   REGION Cyclic Error Checks
       IF NOT #Safety_OK_Delayed THEN //11:1
           "Set_Bit_F"(Bit := 0,
                       Bit_Value := 1,
                       Var := #Cnv_Control.Cnv_Errors.Error_Word_1);
       END_IF;

       IF #Cnv_Control.Motor.Error THEN
           "Set_Bit_F"(Bit := 0,
                       Bit_Value := 1,
                       Var := #Cnv_Control.Cnv_Errors.Error_Word_4);
       END_IF;

       IF #Cnv_Control.Instruction.Stop THEN //HMI STOP
           "Set_Bit_F"(Bit := 1,
                       Bit_Value := 1,
                       Var := #Cnv_Control.Cnv_Errors.Error_Word_1);
       END_IF;

       IF #Cnv_Control.Safety_Stop_Cnrl.Error THEN
           "Set_Bit_F"(Bit := 1,
                       Bit_Value := 1,
                       Var := #Cnv_Control.Cnv_Errors.Error_Word_4);
       END_IF;

       // IF ((#ID_Decoded.VTD = 1 AND "Errors_Profinet_1".%X8) OR
       //     (#ID_Decoded.VTD = 2 AND "Errors_Profinet_3".%X7) OR
       //     (*#ID_Decoded.VTD = 3 AND "Errors_Profinet_5".%X4) OR *)
       //     (#ID_Decoded.VTD = 4 AND "Errors_Profinet_7".%X1) OR
       //     (#ID_Decoded.VTD = 5 AND "Errors_Profinet_8".%X6)) AND #Cnv_Control.Mode <> 1
       // THEN //Profinet error
       //     "Set_Bit_F"(Bit := 3,
       //                 Bit_Value := 1,
       //                 Var := #Cnv_Control.Cnv_Errors.Error_Word_3);
       // END_IF;


       // go to error state
       IF #Cnv_Control.Cnv_Errors.Error_Word_1 <> 0 OR
           #Cnv_Control.Cnv_Errors.Error_Word_2 <> 0 OR
           #Cnv_Control.Cnv_Errors.Error_Word_3 <> 0 OR
           #Cnv_Control.Cnv_Errors.Error_Word_4 <> 0
       THEN
           #Cnv_Control.Error := TRUE;
           #State := 400;
       END_IF;
   END_REGION

   REGION VFD
       //Status
       #Cnv_Control.Motor.Ready := (#Cnv_Control.Inputs.VFD_Status.%X0 OR #Cnv_Control.Inputs.VFD_Status.%X1) AND NOT #Cnv_Control.Motor.Error;
       #Cnv_Control.Motor.Error := #Cnv_Control.Inputs.VFD_Status.%X3 OR #Cnv_Control.Inputs.VFD_Status.%X7 OR NOT #Cnv_Control.Inputs.VFD_Status.%X13;
       #Cnv_Control.Motor.Enabled := #Cnv_Control.Inputs.VFD_Status.%X2;
       #Cnv_Control.Motor.Actual_Current := SCALE_X(MIN := 0,
                                                    VALUE := NORM_X(MIN := 0,
                                                                    VALUE := #Cnv_Control.Inputs.VFD_ActualCurrent,
                                                                    MAX := 16384),
                                                    MAX := 1.98);


       //Actual Speed
       IF #MainSetpoint > 0 THEN
           #Cnv_Control.Motor.Speed_Actual := SCALE_X(MIN := 0,
                                                      VALUE := NORM_X(MIN := 0,
                                                                      VALUE := #Cnv_Control.Inputs.VFD_Speed_Actual,
                                                                      MAX := 16384),
                                                      MAX := 130);

           #Cnv_Control.Motor.Actual_Torque := SCALE_X(MIN := 0,
                                                       VALUE := NORM_X(MIN := 0,
                                                                       VALUE := #Cnv_Control.Inputs.VFD_ActualTorque,
                                                                       MAX := 16384),
                                                       MAX := 100);
       ELSIF #MainSetpoint < 0 THEN
           #Cnv_Control.Motor.Speed_Actual := SCALE_X(MIN := 0,
                                                      VALUE := NORM_X(MIN := 0,
                                                                      VALUE := #Cnv_Control.Inputs.VFD_Speed_Actual * -1,
                                                                      MAX := 16384),
                                                      MAX := 130);

           #Cnv_Control.Motor.Actual_Torque := SCALE_X(MIN := 0,
                                                       VALUE := NORM_X(MIN := 0,
                                                                       VALUE := #Cnv_Control.Inputs.VFD_ActualTorque * -1,
                                                                       MAX := 16384),
                                                       MAX := 100);
       ELSE
           #Cnv_Control.Motor.Speed_Actual := 0;
           #Cnv_Control.Motor.Actual_Torque := 0;
       END_IF;

       //MAIN SETPOINT
       IF #Cnv_Control.Motor.Forward THEN
           #MainSetpoint := (SCALE_X(MIN := 0,
                                     VALUE := NORM_X(MIN := 0,
                                                     VALUE := #Cnv_Control.Motor.Speed (** 1.681*),
                                                     MAX := 130),
                                     MAX := 1865.0) * -1);
       ELSIF #Cnv_Control.Motor.Reverse THEN
           #MainSetpoint := SCALE_X(MIN := 0,
                                    VALUE := NORM_X(MIN := 0,
                                                    VALUE := #Cnv_Control.Motor.Speed (** 1.681*),
                                                    MAX := 130),
                                    MAX := 1865.0);
       ELSE
           #MainSetpoint := 0;
       END_IF;

       IF #Safety_OK THEN
           #ConfigAxis := 16#003F;
       ELSE
           #ConfigAxis := 16#003D;
       END_IF;

           #SinaSpeed(EnableAxis := #Cnv_Control.Motor.Forward OR #Cnv_Control.Motor.Reverse,
                      AckError := #Cnv_Control.Instruction.Reset OR "Reset_All" OR #HMI_Reset,
                      SpeedSp := #MainSetpoint,
                      RefSpeed := 1865.0,
                      ConfigAxis := #ConfigAxis,
                      HWIDSTW := #Cnv_Settings.G120_Hardware_ID,
                      HWIDZSW := #Cnv_Settings.G120_Hardware_ID);


   END_REGION

   #HMI_Reset := "Screen_DB_1".Reset_All[1] OR "Screen_DB_1".Reset_All[2] OR "CNV_HMI"."Reset(1)"[1] OR "CNV_HMI"."Reset(1)"[2];
   ;
END_FUNCTION_BLOCK

FUNCTION_BLOCK "Safety_Stops_FB"   // FB7, SCL
{ S7_Optimized_Access := 'TRUE' }
VERSION : 0.1
// stored: AutoNumber true, IsIECCheckEnabled false, IsRetainMemResEnabled false, MemoryReserve 100, SetENOAutomatically false, UDAEnableTagReadback false
   VAR_INPUT
      Sys_No : UInt;
      Mode : UInt;
      Timeout : UInt;
      Reset : Bool;
   END_VAR
   VAR_IN_OUT
      Sfts_Control : "Sfts_Control";
   END_VAR
   VAR
      State : UInt;
      LP_Timer { ExternalAccessible := 'False'; ExternalVisible := 'False'; ExternalWritable := 'False'} : TON_TIME;
      T_Run { S7_SetPoint := 'True'} : TOF_TIME;
      Timer_1 : Time;
   END_VAR
BEGIN
   #Sfts_Control.Enabled := #Sfts_Control.Instruction.Enable := #Mode = 2 OR #Mode = 3;

   //MODES
   IF (#Mode = 1 OR #Mode = 5) AND NOT #Sfts_Control.Error THEN
       #State := 500;
   END_IF;

   (*
   TODO
   1. Need to add the mode and running checks for manual mode
   2. Add output for safety stop brake.

   Mode select is done via the HMI. Might add external mode select switches.

           Mode select mask:
           0: Disabled
           1: Manual
           2: Semi-Auto
           3: Auto
           4: Teach - N/A for Cnv
           5: Maintenance

   Device ID Format: XXYYZZ    
   XX = Device type   
       01   VTD
       10  Cnv_Front_of_VTD
       11  Cnv_Rear_of_VTD
       12  Cnv_On_Extractor
       20  Safety_Stop_Front_of_VTD
       21  Safety_Stop_Rear_of_VTD
   YY = Floor   
   ZZ = VTD Connected to 
   *)


   REGION Cyclic Checks
       //Update variables
       #Sfts_Control.SM_State := #State;

       #LP_Timer(IN := #Sfts_Control.Running,
                 PT := UINT_TO_TIME(#Timeout));

       //STOPPER STATE
       IF #Sfts_Control.Inputs.DP_Extended AND NOT #Sfts_Control.Inputs.DP_Retracted THEN
           #Sfts_Control.LP_State := 1; // EXTENDED
       ELSIF NOT #Sfts_Control.Inputs.DP_Extended AND #Sfts_Control.Inputs.DP_Retracted THEN
           #Sfts_Control.LP_State := 0; //RETRACTED
       ELSE
           #Sfts_Control.LP_State := 2; //LOST
       END_IF;;
   END_REGION

   REGION Auto Mode 
           CASE #State OF
               0: //IDLE MODE
                   IF #Mode = 2 OR #Mode = 3 THEN
                       IF #Sfts_Control.Instruction.Enable AND #Sfts_Control.Error = 0 THEN
                           #Sfts_Control.Enabled := TRUE;
                           #State := 10;
                       END_IF;
                   END_IF;
               10: //Standby
                   IF NOT #Sfts_Control.Running AND #Sfts_Control.Error = 0 AND
                       (#Sfts_Control.Instruction.Extend AND (#Mode = 3 OR #Mode = 2)) OR (#Sfts_Control.Instruction.Manual_Extend AND #Mode = 2) THEN
                       IF #Sfts_Control.Inputs.DP_Extended THEN
                           ; // Complete the task as the LP ar already extended
                       ELSIF #Sfts_Control.Inputs.DP_Retracted THEN
                           #Sfts_Control.Running := True;
                           #State := 20;
                       ELSE
                           #Sfts_Control.Error := 0; //Unknown locking pin state
                           #State := 400;
                       END_IF;
                   ELSIF NOT #Sfts_Control.Running AND #Sfts_Control.Error = 0 AND
                       (#Sfts_Control.Instruction.Retract AND #Mode = 3) OR (#Sfts_Control.Instruction.Manual_Retract AND #Mode = 2) THEN
                       IF #Sfts_Control.Inputs.DP_Retracted THEN
                           ; // Complete the task as the LP ar already extended
                       ELSIF #Sfts_Control.Inputs.DP_Extended THEN
                           #Sfts_Control.Running := True;
                           #State := 40;
                       ELSE
                           #Sfts_Control.Error := 0; //Unknown locking pin state
                           #State := 400;
                       END_IF;
                   END_IF;

               20: //Extend safety locking pins
                   #Sfts_Control.Motor_Extend := TRUE;
                   IF #Sfts_Control.Inputs.DP_Extended THEN
                       #Sfts_Control.Motor_Extend := FALSE;
                       #Sfts_Control.Running := FALSE;
                       #State := 0;
                   END_IF;

               40: //Retract safety locking pins
                   #Sfts_Control.Motor_Retract := TRUE;
                   IF #Sfts_Control.Inputs.DP_Retracted THEN
                       #Sfts_Control.Motor_Retract := FALSE;
                       #Sfts_Control.Running := FALSE;
                       #State := 0;
                   END_IF;

               400: // Error#Sfts_Control
                   #Sfts_Control.Motor_Retract := FALSE;
                   #Sfts_Control.Motor_Extend := FALSE;
                   #Sfts_Control.Running := FALSE;
                   #LP_Timer(IN := FALSE,
                             PT := T#0S);
                   IF #Reset OR "Reset_All" OR
                       "Screen_DB_1".Reset_All[1] OR "Screen_DB_1".Reset_All[2] OR
                       "CNV_HMI"."Reset(1)"[1] OR "CNV_HMI"."Reset(1)"[2]
                   THEN
                       #Sfts_Control.Error := FALSE;
                       #State := 0;
                   END_IF;

               500:
                   IF #Sfts_Control.Instruction.Manual_Extend AND NOT #Sfts_Control.Inputs.DP_Extended THEN
                       #Sfts_Control.Motor_Extend := TRUE;
                       #Sfts_Control.Running := TRUE;
                   ELSIF #Sfts_Control.Instruction.Manual_Retract AND NOT #Sfts_Control.Inputs.DP_Retracted THEN
                       #Sfts_Control.Motor_Retract := TRUE;
                       #Sfts_Control.Running := TRUE;
                   ELSE
                       #Sfts_Control.Motor_Extend := FALSE;
                       #Sfts_Control.Motor_Retract := FALSE;
                       #Sfts_Control.Running := FALSE;
                   END_IF;

                   IF #Mode <> 1 AND #Mode <> 5 THEN
                       #State := 0;
                   END_IF;
           END_CASE;
   END_REGION

   REGION Cyclic Error Checks
       IF #Sfts_Control.Inputs.DP_Extended AND #Sfts_Control.Inputs.DP_Retracted THEN
           #Sfts_Control.Error := TRUE; //Cant have the locking pins extended and retracted at the same time11
       END_IF;

       // Statement section REGION
       IF #LP_Timer.Q THEN
           #Sfts_Control.Error := TRUE;//locking pin timeout
       END_IF;

       IF #Sfts_Control.Error THEN
           #State := 400;
       END_IF;
   END_REGION

   REGION Assign outputs
       #T_Run(IN := #Sfts_Control.Motor_Extend OR #Sfts_Control.Motor_Retract,
                             PT := #Timer_1);

   END_REGION
END_FUNCTION_BLOCK

FUNCTION_BLOCK "Light_Bars"   // FB6, SCL
{ S7_Optimized_Access := 'TRUE' }
VERSION : 0.1
// stored: AutoNumber true, IsIECCheckEnabled false, IsRetainMemResEnabled false, MemoryReserve 100, SetENOAutomatically false, UDAEnableTagReadback false
   VAR_INPUT
      VTD_Mode : UInt;
      VTD_Speed : Int;
      Fault : Bool;
   END_VAR
   VAR_OUTPUT
      Animation_B1 : Byte;
      Color_B1 : Byte;
      Speed_B1 : Byte;
      Animation_B2 : Byte;
      Color_B2 : Byte;
      Speed_B2 : Byte;
   END_VAR
BEGIN
   //Commands for Light Bar

   IF #VTD_Mode = 0 AND NOT #Fault THEN // (0)Disabled = No light  
       #Animation_B1:= #Animation_B2:= 0;

   ELSIF #VTD_Mode = 1 AND #VTD_Speed = 0 AND  NOT #Fault AND NOT "SinaSpeed_VTD_DB_1".EnableAxis THEN // (1)Manual= Yellow Stop
       #Animation_B1 := #Animation_B2 := 1;
       #Color_B1 := #Color_B2 := 4;

   ELSIF #VTD_Mode = 1 AND #VTD_Speed > 0 AND #VTD_Speed <= 33 AND  NOT #Fault AND "SinaSpeed_VTD_DB_1".EnableAxis THEN // (1)Manual= Yellow until 33%
       #Animation_B1 := #Animation_B2 := 2;
       #Speed_B1 := #Speed_B2 := 2;
       #Color_B1 := #Color_B2 := 4;

   ELSIF #VTD_Mode = 1 AND #VTD_Speed > 33 AND #VTD_Speed <= 100 AND  NOT #Fault THEN // (1)Manual= Yellow until 66%
       #Animation_B1 := #Animation_B2 := 2;
       #Speed_B1 := #Speed_B2 := 0;
       #Color_B1 := #Color_B2 := 4;

   // ELSIF #VTD_Mode = 1 AND #VTD_Speed > 66 AND #VTD_Speed <= 100 AND  NOT #Fault THEN // (1)Manual= Yellow until 100%
   //     #Animation_B1 := #Animation_B2 := 2;
   //     #Speed_B1 := #Speed_B2 := 1;
   //     #Color_B1 := #Color_B2 := 4;

   ELSIF #VTD_Mode = 2 AND #VTD_Speed = 0 AND  NOT #Fault AND NOT "SinaSpeed_VTD_DB_1".EnableAxis THEN // (2)Semi-auto = Blue Stop
       #Animation_B1 := #Animation_B2 := 1;
       #Color_B1 := #Color_B2 := 9;
       #Speed_B1 := #Speed_B2 := 0;

   ELSIF #VTD_Mode = 2 AND #VTD_Speed > 0 AND #VTD_Speed <= 33 AND  NOT #Fault AND "SinaSpeed_VTD_DB_1".EnableAxis THEN // (2)Semi-auto = Blue until 33%
       #Animation_B1 := #Animation_B2 := 2;
       #Speed_B1 := #Speed_B2 := 2;
       #Color_B1 := #Color_B2 := 9;

   ELSIF #VTD_Mode = 2 AND #VTD_Speed > 33 AND #VTD_Speed <= 100 AND  NOT #Fault THEN // (2)Semi-auto = Blue until 66%
       #Animation_B1 := #Animation_B2 := 2;
       #Speed_B1 := #Speed_B2 := 0;
       #Color_B1 := #Color_B2 := 9;

   // ELSIF #VTD_Mode = 2 AND #VTD_Speed > 66 AND #VTD_Speed <= 100 AND  NOT #Fault THEN // (2)Semi-auto = Blue until 100%
   //     #Animation_B1 := #Animation_B2 := 2;
   //     #Speed_B1 := #Speed_B2 := 1;
   //     #Color_B1 := #Color_B2 := 9;

   ELSIF #VTD_Mode = 3 AND #VTD_Speed = 0 AND  NOT #Fault AND NOT "SinaSpeed_VTD_DB_1".EnableAxis THEN // (3)Auto = Green Stop
       #Animation_B1 := #Animation_B2 := 1;
       #Color_B1 := #Color_B2 := 0;

   ELSIF #VTD_Mode = 3 AND #VTD_Speed > 0 AND #VTD_Speed <= 33 AND  NOT #Fault AND "SinaSpeed_VTD_DB_1".EnableAxis THEN // (3)Auto = Green until 33%
       #Animation_B1 := #Animation_B2 := 2;
       #Speed_B1 := #Speed_B2 := 2;
       #Color_B1 := #Color_B2 := 0;

   ELSIF #VTD_Mode = 3 AND #VTD_Speed > 33 AND #VTD_Speed <= 100 AND  NOT #Fault THEN // (3)Auto = Green until 66%
       #Animation_B1 := #Animation_B2 := 2;
       #Speed_B1 := #Speed_B2 := 0;
       #Color_B1 := #Color_B2 := 0;

   // ELSIF #VTD_Mode = 3 AND #VTD_Speed > 66 AND #VTD_Speed <= 100 AND  NOT #Fault THEN // (3)Auto = Green until 100%
   //     #Animation_B1 := #Animation_B2 := 2;
   //     #Speed_B1 := #Speed_B2 := 1;
   //     #Color_B1 := #Color_B2 := 0;

   ELSIF #VTD_Mode = 4 AND #VTD_Speed = 0 AND  NOT #Fault THEN // (4)Tech = Orange Stop
       #Animation_B1 := #Animation_B2 := 1;
       #Color_B1 := #Color_B2 := 2;

   ELSIF #VTD_Mode = 4 AND #VTD_Speed > 0 AND #VTD_Speed <= 33 AND  NOT #Fault THEN // (4)Tech = Orange until 33%
       #Animation_B1 := #Animation_B2 := 2;
       #Speed_B1 := #Speed_B2 := 2;
       #Color_B1 := #Color_B2 := 2;

   ELSIF #VTD_Mode = 4 AND #VTD_Speed > 33 AND #VTD_Speed <= 66 AND  NOT #Fault THEN // (4)Tech = Orange until 66%
       #Animation_B1 := #Animation_B2 := 2;
       #Speed_B1 := #Speed_B2 := 0;
       #Color_B1 := #Color_B2 := 2;

   ELSIF #VTD_Mode = 4 AND #VTD_Speed > 66 AND #VTD_Speed <= 100 AND  NOT #Fault THEN // (4)Tech = Orange until 100%
       #Animation_B1 := #Animation_B2 := 2;
       #Speed_B1 := #Speed_B2 := 1;
       #Color_B1 := #Color_B2 := 2;

   ELSIF #VTD_Mode = 5 AND #VTD_Speed = 0 AND  NOT #Fault THEN // (5)Maintenance = White Stop
       #Animation_B1 := #Animation_B2 := 1;
       #Color_B1 := #Color_B2 := 19;

   ELSIF #VTD_Mode = 5 AND #VTD_Speed > 0 AND #VTD_Speed <= 33 AND  NOT #Fault THEN // (5)Maintenance = White until 33%
       #Animation_B1 := #Animation_B2 := 2;
       #Speed_B1 := #Speed_B2 := 2;
       #Color_B1 := #Color_B2 := 19;

   ELSIF #VTD_Mode = 5 AND #VTD_Speed > 33 AND #VTD_Speed <= 66 AND  NOT #Fault THEN // (5)Maintenance = White until 66%
       #Animation_B1 := #Animation_B2 := 2;
       #Speed_B1 := #Speed_B2 := 0;
       #Color_B1 := #Color_B2 := 19;

   ELSIF #VTD_Mode = 5 AND #VTD_Speed > 66 AND #VTD_Speed <= 100 AND  NOT #Fault THEN // (5)Maintenance = White until 100%
       #Animation_B1 := #Animation_B2 := 2;
       #Speed_B1 := #Speed_B2 := 1;
       #Color_B1 := #Color_B2 := 19;

   ELSIF #Fault THEN // Fault = Flash Red
       #Animation_B1:= #Animation_B2 := 2;
       #Color_B1:=#Color_B2 := 1;
   END_IF;
END_FUNCTION_BLOCK

FUNCTION_BLOCK "SICK_Lector_CLV6xx_PNDP"   // FB72, SCL
TITLE = SICK Lector6xx / CLV6xx function block
{ S7_Optimized_Access := 'TRUE' }
AUTHOR : SICKAG
FAMILY : Ident
VERSION : 1.2
// This function block is used for a communication between a SICK Lector6xx / SICK CLV6xx code reader and a Siemens S7-1200/S7-1500 PLC via  PROFINET/PROFIBUS
// stored: AutoNumber false, IsIECCheckEnabled false, IsRetainMemResEnabled false, MemoryReserve 100, SetENOAutomatically false, UDAEnableTagReadback false
   VAR_INPUT
      HWInputIdent : HW_IO;   // Hardware identification number of the input module
      HWInputLength : USInt;   // Size of the input module
      HWOutputIdent : HW_IO;   // Hardware identification number of the output module
      HWOutputLength : USInt;   // Size of the output module
      CANId : USInt;   // CAN ID (0= Master / No CAN network)
      TOut : Time := T#10s;   // Time out
      Req : Bool;   // A positive edge starts the request
      TriggerOn : Bool;   // Select: Trigger On to open the reading gate via a SW-Trigger command
      TriggerOff : Bool;   // Select: Trigger Off to close the reading gate via a SW-Trigger command
      Matchcode : Bool;   // Select: Matchcode (details at #Data)
      SavePermanent : Bool;   // Select: Save permanent
      ComTest : Bool;   // Select: Communication test
      FreeCommand : Bool;   // Select: Free command (details at #Data)
   END_VAR
   VAR_OUTPUT
      RdDone : Bool;   // Positive edge: A reading result sent by the device was received
      ReqDone : Bool;   // Request done
      ReqBusy : Bool;   // Request in process
      Error : Bool;   // Error detected
      Errorcode : DWord;   // Error code (see documentation)
   END_VAR
   VAR_IN_OUT
      Data : "ST_SICK_Lector_CLV6xx";   // Command arguments and result outputs of the FB actions
   END_VAR
   VAR
      bTriggerReq { ExternalAccessible := 'False'; ExternalVisible := 'False'; ExternalWritable := 'False'} : Bool;   // Rising edge detection
      bTriggerReqMem { ExternalAccessible := 'False'; ExternalVisible := 'False'; ExternalWritable := 'False'} : Bool;   // Rising edge detection
      bTriggerDone { ExternalAccessible := 'False'; ExternalVisible := 'False'; ExternalWritable := 'False'} : Bool;   // Rising edge detection
      bTriggerDoneMem { ExternalAccessible := 'False'; ExternalVisible := 'False'; ExternalWritable := 'False'} : Bool;   // Rising edge detection
      bTriggerError { ExternalAccessible := 'False'; ExternalVisible := 'False'; ExternalWritable := 'False'} : Bool;   // Rising edge detection
      bTriggerErrorMem { ExternalAccessible := 'False'; ExternalVisible := 'False'; ExternalWritable := 'False'} : Bool;   // Rising edge detection
      bCanActive { ExternalAccessible := 'False'; ExternalVisible := 'False'; ExternalWritable := 'False'} : Bool;   // CAN-Bus active flag
      bDeviceState { ExternalAccessible := 'False'; ExternalVisible := 'False'; ExternalWritable := 'False'} : Bool;   // Current device state (True= Edit-Mode | False= Run-Mode)
      bEnforceLogout { ExternalAccessible := 'False'; ExternalVisible := 'False'; ExternalWritable := 'False'} : Bool;   // Logout enforced
      bReqBusyMem : Bool;   // Backup variable
      iStep { ExternalAccessible := 'False'; ExternalVisible := 'False'; ExternalWritable := 'False'} : USInt;   // Currrent FB step
      iCommandIndex { ExternalAccessible := 'False'; ExternalVisible := 'False'; ExternalWritable := 'False'} : Int;   // Command index
      iCommandLength { ExternalAccessible := 'False'; ExternalVisible := 'False'; ExternalWritable := 'False'} : UInt;   // Length of the command that should be send
      iRecordSize { ExternalAccessible := 'False'; ExternalVisible := 'False'; ExternalWritable := 'False'} : UInt;   // Length of the record array
      iCommandSize { ExternalAccessible := 'False'; ExternalVisible := 'False'; ExternalWritable := 'False'} : UInt;   // Length of the command array
      iReadingResultSize { ExternalAccessible := 'False'; ExternalVisible := 'False'; ExternalWritable := 'False'} : UInt;   // Length of the reading result array
      iIndex { ExternalAccessible := 'False'; ExternalVisible := 'False'; ExternalWritable := 'False'} : UInt;   // Index variable
      nTempErrorCode { ExternalAccessible := 'False'; ExternalVisible := 'False'; ExternalWritable := 'False'} : DWord;   // Temporarily error code
      nLogoutErrorCode { ExternalAccessible := 'False'; ExternalVisible := 'False'; ExternalWritable := 'False'} : DWord;   // Temporarily error code
      arrSelection { ExternalAccessible := 'False'; ExternalVisible := 'False'; ExternalWritable := 'False'} : Array[0..5] of Bool;   // input bit selection
      arrCommand { ExternalAccessible := 'False'; ExternalVisible := 'False'; ExternalWritable := 'False'} : Array[0..499] of Byte;   // Contains the transmitted CoLa command
      arrRecord { ExternalAccessible := 'False'; ExternalVisible := 'False'; ExternalWritable := 'False'} : Array[0..499] of Byte;   // Contains the received telegram
      fbTimeout { ExternalAccessible := 'False'; ExternalVisible := 'False'; ExternalWritable := 'False'; S7_SetPoint := 'True'} : TON_TIME;   // Instance: Timer on delay (Time out)
      fbCCom { ExternalAccessible := 'False'; ExternalVisible := 'False'; ExternalWritable := 'False'; S7_SetPoint := 'True'} : "SICK_CCOMM_PNDP";   // Instance: CoLa communication block
   END_VAR
   VAR_TEMP
      iTemp1 : Int;   // Temporarily variable
      iTemp2 : UDInt;   // Temporarily variable
      iTemp3 : UDInt;   // Temporarily variable
      nFncValue : DWord;   // Get/Set function value
      nFncErrorCode : Word;   // Get/Set function error code
   END_VAR
BEGIN
   (*===========================================================================================
   Name:   SICK_Lector_CLV6xx_PNDP 
   Author: SICK AG
   =============================================================================================
   Description: 
   This function block is used for a communication between a SICK Lector6xx / SICK CLV6xx
   code reader and a Siemens S7-1200/S7-1500 PLC via PROFINET/PROFIBUS.                         

   =============================================================================================
   Features:        
   - Receive reading results of the device, triggered by a command, fieldbus or by a hardware 
     switch. The content of the result can be modified in the "Output Format" option in the
     SOPAS engineeringtool.                                           
   - Open and close a reading gate (software trigger via command)
   - Set a new Matchcode evaluation condition 
   - Save all device parameters permanent                                                  
   - Communication test
   - Send a free defined CoLa-A telegram and receive the result
   - All commands can also be used in a SICK CAN-Bus network

   =============================================================================================
   Version history:
   Date       | Version | Author  | Remark
   ---------------------------------------------------------------------------------------------
   21/02/2014 | V1.0    | SICK AG | Initial version
   07/08/2014 | V1.1    | SICK AG | Replace R_TRIG function 
   24/10/2017 | V1.2    | SICK AG | Avoid initialization warnings which occurs using TIA V13 or higher
   ============================================================================================*)

   (*===================================== INITIALISATION =====================================*)
   #iRecordSize:= 500;         (*Length of the arrRecord array*)
   #iCommandSize:= 500;        (*Length of the arrCommand array*)
   #iReadingResultSize:= 200;  (*Length of the reading result array*)

   (*Rising edge detection*)
   #bTriggerReq:= #Req AND NOT #bTriggerReqMem;
   #bTriggerReqMem:= #Req;
   #bTriggerDone:= #fbCCom.ReqDone AND NOT #bTriggerDoneMem;
   #bTriggerDoneMem:= #fbCCom.ReqDone;
   #bTriggerError:= #fbCCom.Error AND NOT #bTriggerErrorMem;
   #bTriggerErrorMem:= #fbCCom.Error;

   (*Reset the read done flag every cycle*)
   #RdDone:= false;


   (*===================================== ERROR HANDLING =====================================*)
   (* bDeviceState  |  bEnforceLogout  |  Action
          FALSE     |      FALSE       |  Errorcode = Errorcode from last plc cycle
          FALSE     |      TRUE        |  Errorcode = Logout error
          TRUE      |      FALSE       |  Enforce "Logout" command
          TRUE      |      TRUE        |  Errorcode = Logout not possible + Reason*)
   IF #nTempErrorCode <>16#0000_0000 THEN

     (*Enfore "Logout" command*)
     IF #bDeviceState AND NOT #bEnforceLogout THEN
       #bEnforceLogout:= true;
       #iCommandIndex:= 11;                  (*Logout*)
       #nLogoutErrorCode:= #nTempErrorCode;  (*Save current error code*)
       #nTempErrorCode:= 16#0000_0000;       (*Clear currenr error variable*)
       #iStep:= 4;                           (*Create command*)

     (*Logout can not be ensured*)
     ELSIF #bDeviceState AND #bEnforceLogout THEN
       #Errorcode.%W1:= #nTempErrorCode.%W0;  
       #Errorcode.%W0:= 16#0017;  (*Error: Logout can not be ensured (please check the device state)*)

     (*Errorcode = Errorcode from the last plc cycle or logout error*)
     ELSE
       #Errorcode:= #nTempErrorCode;
     END_IF;

     (*Update FB status*)
     IF #nTempErrorCode <> 16#0000_0000 THEN
       #ReqDone:= false;
       #ReqBusy:= false;
       #bReqBusyMem:= false;
       #Error:= true;
       #nTempErrorCode:= 16#0000_0000;
       #nLogoutErrorCode:= 16#0000_0000;
       #iStep:= 0;
       RETURN;
     END_IF;
   END_IF;

   (*Time out detection*)
   #fbTimeout(IN:= #bReqBusyMem, PT:= #TOut);
   IF #fbTimeout.Q THEN
     #nTempErrorCode:= 16#0000_0010; (*Error: Time out*)
   END_IF;

   (*Check if a device error is detected: 'sFA XX'*)
   IF #bTriggerDone AND ((NOT #bCanActive AND
     #arrRecord[0] = 's' AND
     #arrRecord[1] = 'F' AND
     #arrRecord[2] = 'A') OR (#bCanActive AND
     #arrRecord[0] = 's' AND
     #arrRecord[12] = 'F' AND
     #arrRecord[13] = 'A')) THEN

     (*Get the position of the error code*)
     IF #bCanActive THEN
       #iIndex:= 15;
     ELSE
       #iIndex:= 4;
     END_IF;

     "SICK_GetValue"(iTelegramLength:= INT_TO_UINT(#fbCCom.ReqLength),
                     iValueLength:= 0,
                     nValue=> #nFncValue,
                     nErrorCode=> #nFncErrorCode,
                     iPosition:= #iIndex,
                     arrData:= #arrRecord);

     IF #nFncErrorCode = 16#0000 THEN
       #nTempErrorCode.%W1:= DWORD_TO_WORD(#nFncValue);
       #nTempErrorCode.%W0:= 16#0011; (*Error: Device error*)
     ELSE
       #nTempErrorCode.%W1:= #nFncErrorCode;
       #nTempErrorCode.%W0:= 16#0012; (*Error: SICK_GetValue error*)      
     END_IF;
   END_IF;

   (*Error detected*)
   IF #nTempErrorCode <>16#0000_0000 THEN
     RETURN;
   END_IF;


   (*================================= START REQUEST (STEP 1) =================================*)
   IF NOT #bReqBusyMem AND #bTriggerReq THEN
     #ReqDone:= false;
     #ReqBusy:= true;
     #bReqBusyMem:= true;
     #Error:= false;
     #Errorcode:= 16#0000_0000;
     #bDeviceState:= false;
     #bEnforceLogout:= false;

     (*Save the current bit selection for the job*)
     #arrSelection[0]:= #TriggerOn;
     #arrSelection[1]:= #TriggerOff;
     #arrSelection[2]:= #Matchcode;
     #arrSelection[3]:= #SavePermanent;
     #arrSelection[4]:= #ComTest;
     #arrSelection[5]:= #FreeCommand;

     (*Check CAN-ID*)
     IF #CANId > 63 THEN
       #nTempErrorCode:= 16#0000_0014; (*Error invalid CAN Id*)  
     ELSIF #CANId = 0 THEN
       #bCanActive:= false;
       #iStep:= 3; (*Check parameter input*)
     ELSE
       #bCanActive:= true;
       #iStep:= 2; (*Add CAN identifier*)
     END_IF;
   END_IF;


   (*=============================== ADD CAN IDENTIFIER (STEP 2) ==============================*)
   IF #iStep =2 THEN
     Strg_TO_Chars(Strg:= 's{ 00 01 ', pChars:= 0, Cnt=> #iIndex, Chars:=#arrCommand);

     "SICK_SetValue"(bAddBlank:= false,
                     nValue:= #CANId,
                     arrData=> #arrCommand,
                     nErrorCode=> #nFncErrorCode,
                     iPosition:= #iIndex);
     IF #nFncErrorCode <> 16#0000 THEN
       #nTempErrorCode.%W1:= #nFncErrorCode;
       #nTempErrorCode.%W0:= 16#0013; (*Error: SICK_SetValue error*)
     ELSE
       #arrCommand[#iIndex]:= '}';
       #iStep:= 3; (*Check parameter input*)
     END_IF;
   END_IF;


   (*============================= CHECK PARAMETER INPUT (STEP 3) =============================*)
   IF #iStep =3 THEN
     #iTemp1:= 0; (*Counts up the active bit selection*)

     (*Command: Trigger On*)
     IF #arrSelection[0] THEN
       #iTemp1:= #iTemp1+1;
       #iCommandIndex:= 0; (*Send a "Trigger On" command*)
     END_IF;

     (*Command: Trigger Off*)
     IF #arrSelection[1] THEN
       #iTemp1:= #iTemp1+1;
       #iCommandIndex:= 1; (*Send a "Trigger Off" command*)
     END_IF;

     (*Command: Matchcode*)
     IF #arrSelection[2] THEN
       #iTemp1:= #iTemp1+1;

       IF #Data.Matchcode.sName = '' THEN
         #nTempErrorCode:= 16#0000_0022; (*Error: Matchcode name is empty*)
       ELSIF #Data.Matchcode.nCodeType <='$20' OR #Data.Matchcode.nCodeType > '$7E' THEN
         #nTempErrorCode:= 16#0000_0023; (*Error: Invalid code type*)
       END_IF;

       #iCommandIndex:= 10; (*Send a "Login" command*)
     END_IF;

     (*Command: Save permanent*)
     IF #arrSelection[3] THEN 
       #iTemp1:= #iTemp1+1;
       #iCommandIndex:= 10; (*Send a "Login" command*)  
     END_IF;

     (*Command: Communication test*)
     IF #arrSelection[4] THEN
       #iTemp1:= #iTemp1+1;
       #iCommandIndex:= 4; (*Send a "Comm Test" command*)
     END_IF;

     (*Command: Free command*)
     IF #arrSelection[5] THEN
       #iTemp1:= #iTemp1+1;

       (*Check length*)
       IF #bCanActive THEN
         #iTemp2:= INT_TO_UDINT(LEN(#Data.FreeCommand.sCommand))+11;
       ELSE
         #iTemp2:= INT_TO_UDINT(LEN(#Data.FreeCommand.sCommand));
       END_IF;

       IF (LEN(#Data.FreeCommand.sCommand) <=0) OR (#iTemp2 > #iCommandSize) THEN
         #nTempErrorCode:= 16#0000_0020; (*Error: Invalid free command length*)
       END_IF;

       #iCommandIndex:= 5; (*Send a "Free Command" command*)
     END_IF;

     (*Check bit sum of the command selection*)
     IF #iTemp1 <>1 THEN
       #nTempErrorCode:= 16#0000_0015; (*Error: More than one or no parameter selected*)   
     END_IF;

     (*Check if a error was detected*)
     IF #nTempErrorCode = 16#0000_0000 THEN
       #iStep:= 4; (*Create CoLa command*)
     END_IF;
   END_IF;


   (*============================== CREATE COLA COMMAND (STEP 4) ==============================*)
   IF #iStep =4 THEN
     CASE #iCommandIndex OF

     (*Create "Trigger On" command*)
     0:  IF #bCanActive THEN
           Strg_TO_Chars(Strg:= 'MN mTCgateon', pChars:= 12, Cnt=> #iTemp3, Chars:=#arrCommand);
           #iCommandLength:= UDINT_TO_UINT(#iTemp3)+12;
         ELSE
           Strg_TO_Chars(Strg:= 'sMN mTCgateon', pChars:= 0, Cnt=> #iTemp3, Chars:=#arrCommand);
           #iCommandLength:= UDINT_TO_UINT(#iTemp3);
         END_IF;
         #iStep:= 5; (*Send command*)

     (*Create "Trigger Off" command*)
     1:  IF #bCanActive THEN
           Strg_TO_Chars(Strg:= 'MN mTCgateoff', pChars:= 12, Cnt=> #iTemp3, Chars:=#arrCommand);
           #iCommandLength:= UDINT_TO_UINT(#iTemp3)+12;
         ELSE
           Strg_TO_Chars(Strg:= 'sMN mTCgateoff', pChars:= 0, Cnt=> #iTemp3, Chars:=#arrCommand);
           #iCommandLength:= UDINT_TO_UINT(#iTemp3);
         END_IF;
         #iStep:= 5; (*Send command*)

     (*Create "Matchcode" command*)
     2:  IF #bCanActive THEN
           Strg_TO_Chars(Strg:= 'MN mEVSetMatchCode 00 ', pChars:= 12, Cnt=> #iTemp3, Chars:=#arrCommand);
           #iIndex:= UDINT_TO_UINT(#iTemp3+12);
         ELSE
           Strg_TO_Chars(Strg:= 'sMN mEVSetMatchCode 00 ', pChars:= 0, Cnt=> #iTemp3, Chars:=#arrCommand);
           #iIndex:= UDINT_TO_UINT(#iTemp3);
         END_IF;

         (*Add matchcode name*)
         Strg_TO_Chars(Strg:= CONCAT(IN1:= 'name="', IN2:= #Data.Matchcode.sName), pChars:= #iIndex, Cnt=> #iTemp3, Chars:=#arrCommand);
         #iIndex:= #iIndex+UDINT_TO_UINT(#iTemp3);

         (*Add codeType*)
         Strg_TO_Chars(Strg:= '" codeType="', pChars:= #iIndex, Cnt=> #iTemp3, Chars:=#arrCommand);
         #iIndex:= #iIndex+UDINT_TO_UINT(#iTemp3);
         IF #Data.Matchcode.nCodeType = '*' THEN
           Strg_TO_Chars(Strg:= 'dontCare', pChars:= #iIndex, Cnt=> #iTemp3, Chars:=#arrCommand);
           #iIndex:= #iIndex+UDINT_TO_UINT(#iTemp3);
         ELSE
           #arrCommand[#iIndex]:= #Data.Matchcode.nCodeType;
           #iIndex:= #iIndex+1;
         END_IF;

         (*Add Min/Max length*)
         Strg_TO_Chars(Strg:= '" length="', pChars:= #iIndex, Cnt=> #iTemp3, Chars:=#arrCommand);
         #iIndex:= #iIndex+UDINT_TO_UINT(#iTemp3);
         IF #Data.Matchcode.iMinMaxLength = 0 THEN
           Strg_TO_Chars(Strg:= 'dontCare', pChars:= #iIndex, Cnt=> #iTemp3, Chars:=#arrCommand);
           #iIndex:= #iIndex+UDINT_TO_UINT(#iTemp3);
         ELSE
           #arrCommand[#iIndex]:= ((#Data.Matchcode.iMinMaxLength/100) MOD 10)+16#30;     
           #arrCommand[#iIndex+1]:= ((#Data.Matchcode.iMinMaxLength/10) MOD 10)+16#30;
           #arrCommand[#iIndex+2]:= (#Data.Matchcode.iMinMaxLength MOD 10)+16#30;
           #iIndex:= #iIndex+3;
         END_IF;

         (*Add content*)
         Strg_TO_Chars(Strg:= CONCAT(IN1:= '" content="', IN2:= #Data.Matchcode.sContent), pChars:= #iIndex, Cnt=> #iTemp3, Chars:=#arrCommand);
         #iIndex:= #iIndex+UDINT_TO_UINT(#iTemp3);
         #arrCommand[#iIndex]:= '"';


         (*Overwrite the matchcode length*)
         IF #bCanActive THEN
           #nFncValue:= #iIndex-33;      (*Length of the #Matchcode command*)
           #iCommandLength:= #iIndex+1;  (*Length of the whole CoLa command*)
           #iIndex:= 31;                 (*Startindex of the matchcode length*)
         ELSE
           #nFncValue:= #iIndex-22;      (*Length of the #Matchcode command*)
           #iCommandLength:= #iIndex+1;  (*Length of the whole CoLa command*)
           #iIndex:= 20;                 (*Startindex of the matchcode length*)
         END_IF;

         "SICK_SetValue"(bAddBlank:= false,
                         nValue:= #nFncValue,
                         arrData=> #arrCommand,
                         nErrorCode=> #nFncErrorCode,
                         iPosition:=#iIndex);
         IF #nFncErrorCode <> 16#0000 THEN
           #nTempErrorCode.%W1:= #nFncErrorCode;
           #nTempErrorCode.%W0:= 16#0013; (*Error: SICK_SetValue error*)
         ELSE
           #iStep:= 5; (*Send command*)
         END_IF;

     (*Create "Save Permanent" command*)   
     3:  IF #bCanActive THEN
           Strg_TO_Chars(Strg:= 'MN mEEwriteall', pChars:= 12, Cnt=> #iTemp3, Chars:=#arrCommand);
           #iCommandLength:= UDINT_TO_UINT(#iTemp3+12);
         ELSE
           Strg_TO_Chars(Strg:= 'sMN mEEwriteall', pChars:= 0, Cnt=> #iTemp3, Chars:=#arrCommand);
           #iCommandLength:= UDINT_TO_UINT(#iTemp3);
         END_IF;
         #iStep:= 5; (*Send command*)

     (*Create "Communication Test" command*)
     4:  IF #bCanActive THEN
           Strg_TO_Chars(Strg:= 'RI0', pChars:= 12, Cnt=> #iTemp3, Chars:=#arrCommand);
           #iCommandLength:= UDINT_TO_UINT(#iTemp3)+12;
         ELSE
           Strg_TO_Chars(Strg:= 'sRI0', pChars:= 0, Cnt=> #iTemp3, Chars:=#arrCommand);
           #iCommandLength:= UDINT_TO_UINT(#iTemp3);
         END_IF;
         #iStep:= 5; (*Send command*)

     (*Create "Free Command"*)
     5:  IF #bCanActive THEN
           Strg_TO_Chars(Strg:= DELETE(IN:= #Data.FreeCommand.sCommand, L:=1, P:=1), pChars:= 12, Cnt=> #iTemp3, Chars:=#arrCommand);
           #iCommandLength:= UDINT_TO_UINT(#iTemp3)+12;
         ELSE
           Strg_TO_Chars(Strg:= #Data.FreeCommand.sCommand, pChars:= 0, Cnt=> #iTemp3, Chars:=#arrCommand);
           #iCommandLength:= UDINT_TO_UINT(#iTemp3);
         END_IF;
         #iStep:= 5; (*Send command*)

     (*Create "Login" command*)
     10: IF #bCanActive THEN
           Strg_TO_Chars(Strg:= 'MN SetAccessMode 03 F4724744', pChars:= 12, Cnt=> #iTemp3, Chars:=#arrCommand);
           #iCommandLength:= UDINT_TO_UINT(#iTemp3)+12;
         ELSE
           Strg_TO_Chars(Strg:= 'sMN SetAccessMode 03 F4724744', pChars:= 0, Cnt=> #iTemp3, Chars:=#arrCommand);
           #iCommandLength:= UDINT_TO_UINT(#iTemp3);
         END_IF;
         #iStep:= 5; (*Send command*)

     (*Create "Logout" command*)
     11: IF #bCanActive THEN
           Strg_TO_Chars(Strg:= 'MN Run', pChars:= 12, Cnt=> #iTemp3, Chars:=#arrCommand);
           #iCommandLength:= UDINT_TO_UINT(#iTemp3)+12;
         ELSE
           Strg_TO_Chars(Strg:= 'sMN Run', pChars:= 0, Cnt=> #iTemp3, Chars:=#arrCommand);
           #iCommandLength:= UDINT_TO_UINT(#iTemp3);
         END_IF;
         #iStep:= 5; (*Send command*)

       END_CASE;
   END_IF;


   (*=============================== SEND COLA COMMAND (STEP 5) ===============================*)
   IF #iStep =5 THEN
     IF NOT #fbCCom.ReqBusy AND NOT #bTriggerDone AND NOT #bTriggerError THEN
       #fbCCom.Req:= true;
       #iStep:= 6; (*Wait for the command answer*)
     END_IF;
   END_IF;


   (*========================== WAIT FOR THE COMMAND ANSWER (STEP 6) ==========================*)
   IF #iStep =6 THEN
     (*Communication error*)
     IF #bTriggerError THEN
       #nTempErrorCode:= #fbCCom.Errorcode; (*Error: Communication error*)

       (*Communication done*)
     ELSIF #bTriggerDone THEN
       #iStep:= 7; (*Check the command answer*)
     END_IF;
   END_IF;


   (*============================= CHECK COMMAND RESPONSE (STEP 7) ============================*)
   IF #iStep =7 THEN
     CASE #iCommandIndex OF

     (*Check "Trigger On" response*)
     0:  IF #bCanActive THEN
           IF #arrRecord[0] = 's' AND
             #arrRecord[12] = 'A' AND
             #arrRecord[13] = 'N' AND
             #arrRecord[22] = 'o' AND
             #arrRecord[23] = 'n' AND
             #arrRecord[24] = ' ' AND
             #arrRecord[25] = '1' THEN

             #iStep:= 8; (*Action performed*)
           ELSE
             #nTempErrorCode:= 16#0000_0016; (*Error: Invalid device answer*)                    
           END_IF;
         ELSE
           IF #arrRecord[0] = 's' AND
             #arrRecord[1] = 'A' AND
             #arrRecord[2] = 'N' AND
             #arrRecord[11] = 'o' AND
             #arrRecord[12] = 'n' AND
             #arrRecord[13] = ' ' AND
             #arrRecord[14] = '1' THEN

             #iStep:= 8; (*Action performed*)
           ELSE
             #nTempErrorCode:= 16#0000_0016; (*Error: Invalid device answer*)        
           END_IF;
         END_IF;

     (*Check "Trigger Off" response*)
     1:  IF #bCanActive THEN
           IF #arrRecord[0] = 's' AND
             #arrRecord[12] = 'A' AND
             #arrRecord[13] = 'N' AND
             #arrRecord[22] = 'o' AND
             #arrRecord[23] = 'f' AND
             #arrRecord[24] = 'f' AND
             #arrRecord[25] = ' ' AND
             #arrRecord[26] = '1' THEN

             #iStep:= 8; (*Action performed*)
           ELSE
             #nTempErrorCode:= 16#0000_0016; (*Error: Invalid device answer*)          
           END_IF;
         ELSE
           IF #arrRecord[0] = 's' AND
             #arrRecord[1] = 'A' AND
             #arrRecord[2] = 'N' AND
             #arrRecord[11] = 'o' AND
             #arrRecord[12] = 'f' AND
             #arrRecord[13] = 'f' AND
             #arrRecord[14] = ' ' AND
             #arrRecord[15] = '1' THEN

             #iStep:= 8; (*Action performed*)
           ELSE  
             #nTempErrorCode:= 16#0000_0016; (*Error: Invalid device answer*)          
           END_IF;
         END_IF;

     (*Check "Matchcode" response*)
     2:  IF #bCanActive THEN
           IF NOT(#arrRecord[0] = 's' AND
             #arrRecord[12] = 'A' AND
             #arrRecord[13] = 'N' AND
             #arrRecord[27] = 'o' AND
             #arrRecord[28] = 'd' AND
             #arrRecord[29] = 'e' AND
             #arrRecord[30] = ' ' AND
             #arrRecord[31] = '1') THEN

             #nTempErrorCode:= 16#0000_0016; (*Error: Invalid device answer*)          
           END_IF;
         ELSE
           IF NOT(#arrRecord[0] = 's' AND
             #arrRecord[1] = 'A' AND
             #arrRecord[2] = 'N' AND
             #arrRecord[16] = 'o' AND
             #arrRecord[17] = 'd' AND
             #arrRecord[18] = 'e' AND
             #arrRecord[19] = ' ' AND
             #arrRecord[20] = '1') THEN

             #nTempErrorCode:= 16#0000_0016; (*Error: Invalid device answer*)          
           END_IF;
         END_IF;

         IF #nTempErrorCode = 0 THEN
           #iCommandIndex:= 11; (*Logout*)
           #iStep:= 4;         (*Create command*)
         END_IF;    

     (*Check "Save Permanent" response*)
     3:  IF #bCanActive THEN
           IF NOT(#arrRecord[0] = 's' AND
             #arrRecord[12] = 'A' AND
             #arrRecord[13] = 'N' AND
             #arrRecord[23] = 'a' AND
             #arrRecord[24] = 'l' AND
             #arrRecord[25] = 'l' AND
             #arrRecord[26] = ' ' AND
             #arrRecord[27] = '1') THEN

             #nTempErrorCode:= 16#0000_0016; (*Error: Invalid device answer*)          
           END_IF;
         ELSE
           IF NOT(#arrRecord[0] = 's' AND
             #arrRecord[1] = 'A' AND
             #arrRecord[2] = 'N' AND
             #arrRecord[12] = 'a' AND
             #arrRecord[13] = 'l' AND
             #arrRecord[14] = 'l' AND
             #arrRecord[15] = ' ' AND
             #arrRecord[16] = '1') THEN

             #nTempErrorCode:= 16#0000_0016; (*Error: Invalid device answer*)          
           END_IF;
         END_IF;

         IF #nTempErrorCode = 0 THEN
           #iCommandIndex:= 11; (*Logout*)
           #iStep:= 4;         (*Create command*)
         END_IF;

     (*Check "Communication Test" response*)
     4:  IF #bCanActive THEN
           IF #arrRecord[0] = 's' AND
             #arrRecord[12] = 'R' AND
             #arrRecord[13] = 'A' AND
             #arrRecord[14] = ' ' THEN

             #iStep:= 8; (*Action performed*)
           ELSE
             #nTempErrorCode:= 16#0000_0016; (*Error: Invalid device answer*)          
           END_IF;
         ELSE
           IF #arrRecord[0] = 's' AND
             #arrRecord[1] = 'R' AND
             #arrRecord[2] = 'A' AND
             #arrRecord[3] = ' ' THEN

             #iStep:= 8; (*Action performed*)
           ELSE  
             #nTempErrorCode:= 16#0000_0016; (*Error: Invalid device answer*)          
           END_IF;
         END_IF;

     (*Check "Free command" response*)
     5:  IF #fbCCom.ReqLength <= MAX_LEN(#Data.FreeCommand.sResult) THEN 
           Chars_TO_Strg(Chars:= #arrRecord, pChars:= 0, Cnt:= INT_TO_UINT(#fbCCom.ReqLength),Strg=> #Data.FreeCommand.sResult);
           #iStep:= 8; (*Action performed*)
         ELSE
           #nTempErrorCode:= 16#0000_0021; (*Error: Free command result > Result string*)
         END_IF;

     (*Check "Login" response*)
     10:  IF #bCanActive THEN
           IF NOT(#arrRecord[0] = 's' AND
             #arrRecord[12] = 'A' AND
             #arrRecord[13] = 'N' AND
             #arrRecord[24] = 'M' AND
             #arrRecord[25] = 'o' AND
             #arrRecord[26] = 'd' AND
             #arrRecord[27] = 'e' AND
             #arrRecord[28] = ' ' AND
             #arrRecord[29] = '1') THEN

             #nTempErrorCode:= 16#0000_0016; (*Error: Invalid device answer*)          
           END_IF;
         ELSE
           IF NOT(#arrRecord[0] = 's' AND
             #arrRecord[1] = 'A' AND
             #arrRecord[2] = 'N' AND
             #arrRecord[13] = 'M' AND
             #arrRecord[14] = 'o' AND
             #arrRecord[15] = 'd' AND
             #arrRecord[16] = 'e' AND
             #arrRecord[17] = ' ' AND
             #arrRecord[18] = '1') THEN

             #nTempErrorCode:= 16#0000_0016; (*Error: Invalid device answer*)          
           END_IF;
         END_IF;

         IF #nTempErrorCode = 0 THEN
           IF #arrSelection[2] THEN
             #iCommandIndex:= 2; (*Matchcode*)
             #iStep:= 4;         (*Create command*)
           ELSIF #arrSelection[3] THEN
             #iCommandIndex:= 3; (*Save permanent*)
             #iStep:= 4;         (*Create command*)       
           END_IF;
           #bDeviceState:= true; (*Edit-Mode active*)
         END_IF;

     (*Check "Logout" response*)
     11:  IF #bCanActive THEN
           IF #arrRecord[0] = 's' AND
             #arrRecord[12] = 'A' AND
             #arrRecord[13] = 'N' AND
             #arrRecord[14] = ' ' AND
             #arrRecord[15] = 'R' AND
             #arrRecord[16] = 'u' AND
             #arrRecord[17] = 'n' AND
             #arrRecord[18] = ' ' AND
             #arrRecord[19] = '1' THEN

             #bDeviceState:= false; (*Run-Mode active*)
             #iStep:= 8; (*Action performed*)
           ELSE
             #nTempErrorCode:= 16#0000_0016; (*Error: Invalid device answer*)          
           END_IF;
         ELSE
           IF #arrRecord[0] = 's' AND
             #arrRecord[1] = 'A' AND
             #arrRecord[2] = 'N' AND
             #arrRecord[3] = ' ' AND
             #arrRecord[4] = 'R' AND
             #arrRecord[5] = 'u' AND
             #arrRecord[6] = 'n' AND
             #arrRecord[7] = ' ' AND
             #arrRecord[8] = '1' THEN

             #bDeviceState:= false; (*Run-Mode active*)
             #iStep:= 8; (*Action performed*)
           ELSE  
             #nTempErrorCode:= 16#0000_0016; (*Error: Invalid device answer*)          
           END_IF;
         END_IF;
     END_CASE;
   END_IF;


   (*================================ ACTION PERFORMED (STEP 8) ===============================*)
   IF #iStep =8 THEN
     IF #bEnforceLogout THEN
       #nTempErrorCode:= #nLogoutErrorCode;
     ELSE
       #ReqDone:= true;
       #ReqBusy:= false;
       #bReqBusyMem:= false;
       #iStep:= 0;
     END_IF;
   END_IF;


   (*====================================== COMMUNICATION =====================================*)
   #fbCCom(HWInputIdent:= #HWInputIdent,
           HWInputLength:= #HWInputLength,
           HWOutputIdent:= #HWOutputIdent,
           HWOutputLength:= #HWOutputLength,
           TOut:= #TOut+T#1s,
           CommandLength:= #iCommandLength,
           arrCommand:= #arrCommand,
           arrRecord:= #arrRecord);

   (*Reset the request flag every cycle*)
   #fbCCom.Req:= false;

   (*Read result error*)
   IF #fbCCom.RdLength <0 AND #fbCCom.RdDone THEN
     #Data.ReadingResult.iLength:= -1; (*Error: Reading result longer than record array*)
     FOR #iTemp1:= 1 TO UINT_TO_INT(#iReadingResultSize) DO
       #Data.ReadingResult.arrResult[#iTemp1]:= 16#00;
     END_FOR;

   (*Handling of the reading result*)
   ELSIF #fbCCom.RdDone THEN
     IF #fbCCom.RdLength > #iReadingResultSize THEN
       #Data.ReadingResult.iLength:= -1; (*Error: Reading result longer than reading result array*)
       FOR #iTemp1:= 1 TO UINT_TO_INT(#iReadingResultSize) DO
         #Data.ReadingResult.arrResult[#iTemp1]:= 16#00;
       END_FOR;
     ELSE
       MOVE_BLK(IN:= #arrRecord[0], COUNT:= INT_TO_UINT(#fbCCom.RdLength), OUT=> #Data.ReadingResult.arrResult[1]);
       IF (#Data.ReadingResult.iCounter >=255) THEN
         #Data.ReadingResult.iCounter:= 0;
       ELSE
         #Data.ReadingResult.iCounter:= #Data.ReadingResult.iCounter+1;
       END_IF;
       #Data.ReadingResult.iLength:= #fbCCom.RdLength;
       #RdDone:= true;
     END_IF;
   END_IF;
END_FUNCTION_BLOCK

FUNCTION_BLOCK "SICK_CCOMM_PNDP"   // FB10, SCL
TITLE = SICK_CCOM_PNDP
{ S7_Optimized_Access := 'TRUE' }
AUTHOR : SICKAG
FAMILY : Ident
VERSION : 1.2
// The function block use a Profinet/Probibus connection to communicate with a SICK AutoIdent
// device. The FB makes it possible to send and receive sensor data. The Confirmed Messaging 
// protocol (CM-Protocol) is used to receive even long fragmented read results.
// stored: AutoNumber false, IsIECCheckEnabled false, IsRetainMemResEnabled false, MemoryReserve 100, SetENOAutomatically false, UDAEnableTagReadback false
   VAR_INPUT
      HWInputIdent : HW_IO;   // Hardware identification number of the input module
      HWInputLength : USInt;   // Size of the input module
      HWOutputIdent : HW_IO;   // Hardware identification number of the output module
      HWOutputLength : USInt;   // Size of the output module
      TOut : Time := T#5s;   // Time out
      Req : Bool;   // A positive edge starts the request
      CommandLength : UInt;   // Byte length of the command
   END_VAR
   VAR_OUTPUT
      RdDone : Bool;   // Reading result arrived
      RdLength : Int;   // Byte length of the reading result
      ReqDone : Bool;   // Requested data available
      ReqBusy : Bool;   // Request busy
      ReqLength : Int;   // Byte length of the requested data
      Error : Bool;   // Error
      Errorcode : DWord;   // Error code
   END_VAR
   VAR_IN_OUT
      arrCommand : Array[0..499] of Byte;
      arrRecord : Array[0..499] of Byte;
   END_VAR
   VAR
      bTriggerReq { ExternalAccessible := 'False'; ExternalVisible := 'False'; ExternalWritable := 'False'} : Bool := false;   // Rising edge detection
      bTriggerReqMem { ExternalAccessible := 'False'; ExternalVisible := 'False'; ExternalWritable := 'False'} : Bool := false;   // Rising edge detection
      bReadFrag { ExternalAccessible := 'False'; ExternalVisible := 'False'; ExternalWritable := 'False'} : Bool;
      bWriteFrag { ExternalAccessible := 'False'; ExternalVisible := 'False'; ExternalWritable := 'False'} : Bool;
      bReqBusyMem : Bool;
      iReadStep { ExternalAccessible := 'False'; ExternalVisible := 'False'; ExternalWritable := 'False'} : USInt;
      iWriteStep { ExternalAccessible := 'False'; ExternalVisible := 'False'; ExternalWritable := 'False'} : USInt;
      iReadIndex { ExternalAccessible := 'False'; ExternalVisible := 'False'; ExternalWritable := 'False'} : UInt;
      iWriteIndex { ExternalAccessible := 'False'; ExternalVisible := 'False'; ExternalWritable := 'False'} : UInt;
      iReadHeaderLength { ExternalAccessible := 'False'; ExternalVisible := 'False'; ExternalWritable := 'False'} : UInt;
      iWriteHeaderLength { ExternalAccessible := 'False'; ExternalVisible := 'False'; ExternalWritable := 'False'} : UInt;
      iReadFragmentLength { ExternalAccessible := 'False'; ExternalVisible := 'False'; ExternalWritable := 'False'} : UInt;
      iWriteFragmentLength { ExternalAccessible := 'False'; ExternalVisible := 'False'; ExternalWritable := 'False'} : UInt;
      iRecordSize { ExternalAccessible := 'False'; ExternalVisible := 'False'; ExternalWritable := 'False'} : UInt;
      iCommandSize { ExternalAccessible := 'False'; ExternalVisible := 'False'; ExternalWritable := 'False'} : UInt;
      nTempErrorCode { ExternalAccessible := 'False'; ExternalVisible := 'False'; ExternalWritable := 'False'} : DWord;
      arrInputImage : Array[0..127] of Byte;
      arrOutputImage : Array[0..127] of Byte;
      fbTimeout { ExternalAccessible := 'False'; ExternalVisible := 'False'; ExternalWritable := 'False'; S7_SetPoint := 'True'} : TON_TIME;
   END_VAR
   VAR_TEMP
      iTemp1 : Int;
      iTemp2 : UDInt;
      iTemp3 : UDInt;
   END_VAR
BEGIN
   (*===========================================================================================
   Name:   SICK_CCOMM_PNDP
   Author: SICK AG
   =============================================================================================
   Description: 
   The function block use a Profinet/Probibus connection to communicate with a SICK AutoIdent
   device. The FB makes it possible to send and receive sensor data. The Confirmed Messaging 
   protocol (CM-Protocol) is used to receive even long fragmented read results.

   Send a command:
   The "Req" parameter must be triggered with a rising edge (signal change FALSE to TRUE) in 
   order to carry out the function. For the time during which a valid response has yet to be 
   received from the device, the "ReqBusy" parameter is used to signal  that a response is still 
   pending. The module signals the "ReqDone" = TRUE output parameter when the function has been 
   successfully completed. If data was requested by the device, this data is copied into the 
   Record (arrRecord). The "ReqDone" indicates that new data has been received  for a PLC cycle.
   Only one CoLa-A command request can be send to the same device at one time. 

   Receive a reading result:
   Data sent via trigger command or directly by the device (e.g., direct trigger via a light 
   barrier) is stored in the Record (arrRecord). The "RdDone" output indicates that new data 
   has been received for a PLC cycle. The data sent by the device can be changed or adapted in 
   output format of SOPAS-ET. 

   This AOI supports the folowing SICK devices:
   - Lector6xx
   - RFU6xx
   - CLV6xx 
   - RFH6xx
   =============================================================================================
   Confirmed Messaging Protocol definitions:
   arrInputImage[0]        = Status byte 
   arrInputImage[1]        = Receive counter
   arrInputImage[2]        = Transmit counter back
   arrInputImage[3]        = Command length LSB
   arrInputImage[4]        = Command length MSB
   arrInputImage[5..127]   = Device response (CoLa-A)

   arrOutputImage[0]       = Status byte 
   arrOutputImage[1]       = Receive counter back
   arrOutputImage[2]       = Transmit counter
   arrOutputImage[3]       = Command length LSB
   arrOutputImage[4]       = Command length MSB
   arrOutputImage[5..127]  = Device request (CoLa-A)
   =============================================================================================
   Version history:
   Date       | Version | Created under               | Author  | Remark
   ---------------------------------------------------------------------------------------------
   16/01/2014 | V1.0    | TIA Portal V12 SP1 Update 2 | SICK AG | Initial version
   07/08/2014 | V1.1    | TIA Portal V12 SP1 Update 4 | SICK AG | Replace R_TRIG function 
   22/04/2015 | V1.2    | TIA Portal V12 SP1 Update 4 | SICK AG | Avoid warnings that occur with 
                                                                  TIA V13
   ============================================================================================*)

   (*===================================== INITIALISATION =====================================*)
   #iRecordSize:= 500;   (*Length of the arrRecord array*)
   #iCommandSize:= 500;  (*Length of the arrCommand array*)

   #RdDone:= false;
   #iReadStep:= 0;

   (*Rising edge detection of the request flag*)
   #bTriggerReq:= #Req AND NOT #bTriggerReqMem;
   #bTriggerReqMem:= #Req;

   (*Error detection*)
   IF #nTempErrorCode <>16#0000_0000 THEN
     #ReqDone:= false;
     #ReqBusy:= false;
     #bReqBusyMem:= false;
     #Error:= true;
     #Errorcode:= #nTempErrorCode;
     #nTempErrorCode:= 16#0000_0000;
     #ReqLength:= 0;
     #iWriteStep:= 0;
     RETURN;
   END_IF;

   (*Time out detection*)
   #fbTimeout(IN:=#bReqBusyMem, PT:=#TOut);
   IF #fbTimeout.Q THEN
     #nTempErrorCode:= 16#0000_0001; (*Error: Time out*) 
   END_IF;

   (*Check the hardware ident length of the input module*)
   IF #HWInputLength <8 OR #HWInputLength >128 THEN
     #nTempErrorCode:= 16#0000_0002; (*Error: Incorrect module input length*)
   END_IF;

   (*Check the hardware ident length of the output module*)
   IF #HWOutputLength <8 OR #HWOutputLength >128 THEN
     #nTempErrorCode:= 16#0000_0003; (*Error: Incorrect module output length*)
   END_IF;

   (*Error detected*)
   IF #nTempErrorCode <>16#0000_0000 THEN
     RETURN;
   END_IF;


   (*===================================== COMMUNICATION ======================================*)
   (*Set output data*)
   #iTemp1:= DPWR_DAT(LADDR:= #HWOutputIdent, RECORD:= #arrOutputImage);
   IF #iTemp1 <>0 THEN
     #nTempErrorCode.%W1:= #iTemp1;
     #nTempErrorCode.%W0:= 16#0004; (*Error: Set output data via DPWR_DAT*)
     RETURN;
   END_IF;

   (*Get input data*)
   #iTemp1:= DPRD_DAT(LADDR:= #HWInputIdent, RECORD=> #arrInputImage);
   IF #iTemp1 <>0 THEN
     #nTempErrorCode.%W1:= #iTemp1;
     #nTempErrorCode.%W0:= 16#0005; (*Error: Get input data via DPRD_DAT*)
     RETURN;
   END_IF;

   (*Receive counter ==0 && Receive counter back <>0*)
   IF #arrInputImage[1] =0 AND #arrOutputImage[1] <>0 THEN
     #arrOutputImage[1]:= #arrInputImage[1]; (*Recive counter => Receive counter back*)
     RETURN;
   END_IF;

   (*Transmit counter <> Transmit counter back*)
   IF NOT #bReqBusyMem AND (#arrInputImage[2] <> #arrOutputImage[2]) THEN
     #arrOutputImage[2]:= 0; (*0 => Transmit counter*)
     RETURN;
   END_IF;


   (*============================== HANDLING OF THE RECEIVED DATA =============================*)
   (*New telegram available*)
   IF NOT (#arrInputImage[1] = #arrOutputImage[1]) THEN

     (*Reset error every incoming telegram (Read only mode, e.g. for hand held scanners)*)
     IF #CommandLength <=0 THEN
       #Error:= false;
       #Errorcode:= 16#0000_0000;
     END_IF;

     (*Confirm the receive counter*)
     #arrOutputImage[1]:= #arrInputImage[1];

     (*Get telegram length from the received header*)
     #iReadHeaderLength.%B0:= #arrInputImage[3];
     #iReadHeaderLength.%B1:= #arrInputImage[4];

     (*Check if fragmentation is not active at the moment*)
     IF NOT #bReadFrag THEN
       #iReadIndex:= 0;

       (*Check if fragmentation is needed*)
       IF (#HWInputLength-5) < #iReadHeaderLength THEN
         #bReadFrag:= true;
       END_IF;
     END_IF;

     (*Fragmentation is needed*)
     IF #bReadFrag THEN
       IF (#HWInputLength-5) < #iReadHeaderLength THEN
         #iReadFragmentLength:= #HWInputLength-5;
       ELSE
         #iReadFragmentLength:= #iReadHeaderLength;
       END_IF;

     (*No fragmentation needed*)
     ELSE
       #iReadFragmentLength:= #iReadHeaderLength;
     END_IF;

     (*Copy input data into the output record*)
     IF (#iReadIndex+#iReadFragmentLength) <= #iRecordSize THEN
       MOVE_BLK(IN:= #arrInputImage[5], COUNT:= #iReadFragmentLength, OUT=> #arrRecord[#iReadIndex]);
     END_IF;

     (*Check if all data has been received*)
     IF (#HWInputLength-5) < #iReadHeaderLength THEN
       #iReadIndex:= #iReadIndex+#iReadFragmentLength;

     (*All data has been received*)
     ELSE
       #bReadFrag:= false;
       #iReadStep:= 1;
     END_IF;

     (*Incoming data filter*)
     (* - Check if the receiving telegram os a CoLa answer on a requested 
          comand or a reading result.

         sRA  sWA  sMA  sAN  sAI  sEA  sPX  s{   sSI  sSN  sFA
     sRN  X                                       X    X    X
     sRI  X                                       X    X    X
     sWN       X                                  X    X    X
     sWI       X                                  X    X    X
     sMN            X    X                        X    X    X
     sMI            X         X                   X    X    X
     sEN                           X              X    X    X
     sEI                           X              X    X    X
     sPE                                X         X    X    X
     s{                                      X    X    X    X
     *)
     IF #iReadStep =1 THEN
       (*Filter is only active, while requested data expected*)
       IF #bReqBusyMem THEN
         IF #CommandLength >3 THEN
           (*Get the prefix from the requested command (e.g. 'sRN '*)   
           #iTemp2.%B3:= #arrCommand[0];
           #iTemp2.%B2:= #arrCommand[1];
           #iTemp2.%B1:= #arrCommand[2];
           #iTemp2.%B0:= 16#20;

           (*Get the prefix from the command response (e.g. 'sRA ')*)
           #iTemp3.%B3:= #arrRecord[0];
           #iTemp3.%B2:= #arrRecord[1];
           #iTemp3.%B1:= #arrRecord[2];
           #iTemp3.%B0:= 16#20;
         ELSE
           #iTemp2:= 16#0000_0000;
           #iTemp3:= 16#0000_0000;
         END_IF;

         CASE #iTemp3 OF
         (*'s{  '*)
         16#737B2020:  IF #iTemp2 = 16#737B2020 THEN
                         #iReadStep:= 2; (*Command response*)
                       ELSE
                         #iReadStep:= 3; (*Reading result*)
                       END_IF;

         (*'sRA '*)
         16#73524120:  IF (#iTemp2 = 16#73524E20) OR (#iTemp2 = 16#73524920) THEN
                         #iReadStep:= 2; (*Command response*)
                       ELSE
                         #iReadStep:= 3; (*Reading result*)
                       END_IF;

         (*'sWA '*)
         16#73574120:  IF (#iTemp2 = 16#73574E20) OR (#iTemp2 = 16#73574920) THEN
                         #iReadStep:= 2; (*Command response*)
                       ELSE
                         #iReadStep:= 3; (*Reading result*)
                       END_IF;

         (*'sMA '*)
         16#734D4120:  IF (#iTemp2 = 16#734D4E20) OR (#iTemp2 = 16#734D4920) THEN
                         #iReadStep:= 2; (*Command response*)
                       ELSE
                         #iReadStep:= 3; (*Reading result*)
                       END_IF;

         (*'sAN '*)
         16#73414E20:  IF #iTemp2 = 16#734D4E20 THEN
                         #iReadStep:= 2; (*Command response*)
                       ELSE
                         #iReadStep:= 3; (*Reading result*)
                       END_IF;

         (*'sAI '*)
         16#73414920:  IF #iTemp2 = 16#734D4920 THEN
                         #iReadStep:= 2; (*Command response*)
                       ELSE
                         #iReadStep:= 3; (*Reading result*)
                       END_IF;

         (*'sEA '*)
         16#73454120:  IF (#iTemp2 = 16#73454E20) OR (#iTemp2 = 16#73454920) THEN
                         #iReadStep:= 2; (*Command response*)
                       ELSE
                         #iReadStep:= 3; (*Reading result*)
                       END_IF;

         (*'sPX '*)
         16#73505820:  IF #iTemp2 = 16#73504520 THEN
                         #iReadStep:= 2; (*Command response*)
                       ELSE
                         #iReadStep:= 3; (*Reading result*)
                       END_IF;

         (*'sSI '*)
         16#73534920:  #iReadStep:= 3; (*Reading result*)

         (*'sSN '*)
         16#73534E20:  #iReadStep:= 3; (*Reading result*)

         (*'sFA '*)
         16#73464120:  #iReadStep:= 2; (*Command response*)

         (*Invalid CoLa-A answer*)
         ELSE
           (*Check if a user defined command is used (Request == Response)*)
           FOR #iTemp1:= 0 TO UINT_TO_INT(#CommandLength-1) DO
             IF #arrCommand[#iTemp1] = #arrRecord[#iTemp1] THEN
               #iReadStep:= 2; (*Command response*)
             ELSE
               #iReadStep:= 3; (*Reading result*)
               EXIT;
             END_IF;
           END_FOR;
         END_CASE;

       (*Reading result*)
       ELSE
         #iReadStep:= 3;  (*Reading result*)
       END_IF;
     END_IF;

     (*Incoming telegram is a command response*)
     IF #iReadStep =2 THEN
       IF (#iReadIndex+#iReadFragmentLength) <= #iRecordSize THEN
         #ReqLength:= UDINT_TO_INT(#iReadIndex+#iReadFragmentLength);
         #ReqDone:= true;
         #ReqBusy:= false;
         #bReqBusyMem:= false;
       ELSE
         #nTempErrorCode:= 16#0000_0006; (*Error: Incoming command response > Record size*)
       END_IF;
     END_IF;

     (*Incoming telegram is a reading result*)
     IF #iReadStep =3 THEN
       IF (#iReadIndex+#iReadFragmentLength) <= #iRecordSize THEN
         #RdLength:= UDINT_TO_INT(#iReadIndex+#iReadFragmentLength);
         #RdDone:= true;
       ELSE
         #RdLength:= -1;
         #RdDone:= false;    
       END_IF;
     END_IF;
   END_IF;


   (*=========================== HANDLING OF THE DATA TO BE WRITTEN ===========================*)
   IF #bTriggerReq AND NOT #bReqBusyMem THEN
     #ReqDone:= false;
     #ReqBusy:= true;
     #bReqBusyMem:= true;
     #Error:= false;
     #Errorcode:= 16#0000_0000;
     #iWriteIndex:= 0;

     (*Check command length*)
     IF #CommandLength <=0 THEN
       #nTempErrorCode:= 16#0000_0007; (*Error: Command length <= 0*)
       RETURN;
     ELSIF #CommandLength > #iCommandSize THEN
       #nTempErrorCode:= 16#0000_0008; (*Error: Command length > command array*)
       RETURN;
     END_IF;

     (*Check if the the command telegram must be fragmented*)
     IF (#HWOutputLength-5) < #CommandLength THEN
       #iWriteFragmentLength:= #HWOutputLength-5;
     ELSE
       #iWriteFragmentLength:= #CommandLength;
     END_IF;

     #iWriteHeaderLength:= #CommandLength;
     #iWriteStep:= 1;  
   END_IF;

   (*Write step 1: Command transfer*)
   IF (#iWriteStep =1) AND(#arrInputImage[2] = #arrOutputImage[2]) THEN

     (*Copy command data into the output record*)
     IF((#iWriteIndex+#iWriteFragmentLength) <= #iCommandSize) AND (#iWriteFragmentLength <= (#HWOutputLength-5)) THEN
       MOVE_BLK(IN:= #arrCommand[#iWriteIndex], COUNT:= #iWriteFragmentLength, OUT=> #arrOutputImage[5]);
       (*Increment transmit counter*)
       IF #arrOutputImage[2] = 16#FF THEN
         #arrOutputImage[2]:= 16#01; (*Counter overflow, zero is skipped*)
       ELSE
         #arrOutputImage[2]:= #arrOutputImage[2]+1;
       END_IF;

       (*Set command/fragment length*)
       #arrOutputImage[3]:= #iWriteHeaderLength.%B0;
       #arrOutputImage[4]:= #iWriteHeaderLength.%B1;

       (*Next step*)
       #iWriteStep:= 2;
     ELSE
       #nTempErrorCode:= 16#0000_0009; (*Error: Fragmentation error*)
     END_IF;
       RETURN;
   END_IF;

   (*Write step 2: Fragmentation handling*)
   IF #iWriteStep =2 THEN

     (*Fragmentation is needed*)
     IF (#HWOutputLength-5) < #iWriteHeaderLength THEN
       #bWriteFrag:= true;

       (*Next index*)
       #iWriteIndex:= #iWriteIndex+#iWriteFragmentLength;

       (*Set next header length*)
       #iWriteHeaderLength:= #iWriteHeaderLength-#iWriteFragmentLength;

       (*Set next fragment length*)
       IF (#HWOutputLength-5) < #iWriteHeaderLength THEN
         #iWriteFragmentLength:= #HWOutputLength-5;
       ELSE
         #iWriteFragmentLength:= #iWriteHeaderLength;
       END_IF;

     (*Fragmentation is not needed*)
     ELSE
       #bWriteFrag:= false;
     END_IF;

     (*Next step*)
     #iWriteStep:= 3;
   END_IF;

   (*Write step 3: Check if the transmission of the command/fragment is done*)
   IF #iWriteStep =3 THEN

     (*Transmit counter back == Transmit counter*)
     IF #arrInputImage[2] = #arrOutputImage[2] THEN
       IF #bWriteFrag THEN
         #iWriteStep:= 1;
       ELSE
         #iWriteStep:= 0;
       END_IF;
     END_IF;
   END_IF;
END_FUNCTION_BLOCK

FUNCTION_BLOCK "SICK_Lector_Control_FB"   // FB19, SCL
{ S7_Optimized_Access := 'TRUE' }
VERSION : 0.1
// stored: AutoNumber true, IsIECCheckEnabled false, IsRetainMemResEnabled false, MemoryReserve 100, SetENOAutomatically false, UDAEnableTagReadback false
   VAR_INPUT
      Rd_Done : Bool;
      Req_Done : Bool;
      Req_Busy : Bool;
      Error : Bool;
      arrResult : Array[1..200] of Byte;
      iCounter : USInt;
      iLength : Int;
      Error_Code : DWord;
   END_VAR
   VAR_OUTPUT
      Test_Comm : Bool;
      Enable_Trigger : Bool;
      Disable_Trigger : Bool;
      Enable_Req : Bool;
      Result : String;
      Test_OK : Bool;
   END_VAR
   VAR_IN_OUT
      Test_Comm_HMI : Bool;
      Enable_HMI : Bool;
      Disable_HMI : Bool;
      Auto_Start_Lector : Bool;
      Auto_Stop_Lector : Bool;
   END_VAR
   VAR
      "Timer" { S7_SetPoint := 'True'} : TON_TIME;
      R_Done_DB { S7_SetPoint := 'True'} : R_TRIG;
      T_Reset_DB { S7_SetPoint := 'True'} : TON_TIME;
   END_VAR
BEGIN
   //Communication Test
   IF #Test_Comm_HMI THEN
       #Test_Comm := 1;
       #Enable_Req := 1;
       #Timer.TON(IN:=True,
                              PT:=t#1s);
   END_IF;

   //TEST OK
   IF #Req_Done AND #Timer.Q AND NOT #Error THEN
       #Test_OK := 1;
       #Test_Comm := 0;
       #Enable_Req := 0;
       #Test_Comm_HMI := 0;
       #Timer.TON(IN := FALSE,
                              PT := t#0s);
   END_IF;

   //ERROR
   IF #Timer.Q AND #Error THEN
           #Test_OK := 0;
           #Test_Comm := 0;
           #Enable_Req := 0;
           #Test_Comm_HMI := 0;
           #Timer.TON(IN := FALSE,
                                  PT := t#0s);
       END_IF;

   //Enable Trigger
       IF #Enable_HMI OR #Auto_Start_Lector THEN
       #Enable_Trigger := 1;
       #Enable_Req := 1;
       #Disable_HMI := 0;
       #Disable_Trigger := 0;
   //Disable Trigger
   ELSIF #Disable_HMI OR #"Auto_Stop_Lector" THEN
       #Disable_Trigger := 1;
       #Enable_Req := 1;
       #Enable_HMI := 0;
       #Enable_Trigger := 0;
   ELSE
       #Enable_Trigger := 0;
       #Enable_Req := 0;
       #Disable_Trigger := 0;
   END_IF;


   #R_Done_DB(CLK:=#Rd_Done);

   IF #R_Done_DB.Q OR #T_Reset_DB.Q OR
       (#Enable_HMI AND #Disable_HMI)
   THEN
       #Disable_HMI := 0;
       #Enable_Trigger := 0;
       #Disable_Trigger := 0;
       #Enable_Req := 0;
       #T_Reset_DB.TON(IN := FALSE,
                               PT := T#0S);
               #Auto_Stop_Lector := 0;
   END_IF;

   #T_Reset_DB(IN:=(#Enable_HMI OR #Disable_HMI OR #Auto_Start_Lector OR #Auto_Stop_Lector),
                 PT:=T#10S);


   #Result := "ByteArrayToString_1"(Lenght := #iLength, ByteArray := #arrResult);
END_FUNCTION_BLOCK

FUNCTION_BLOCK "Barcode_Station_FB"   // FB33, SCL
{ S7_Optimized_Access := 'TRUE' }
VERSION : 0.1
// stored: AutoNumber true, IsIECCheckEnabled false, IsRetainMemResEnabled false, MemoryReserve 100, SetENOAutomatically false, UDAEnableTagReadback false
   VAR_INPUT
      Sick_Result : String;
   END_VAR
   VAR_OUTPUT
      "Counter" : UInt;
   END_VAR
   VAR_IN_OUT
      Station_Control : "Barcode_Station_UDT";
      Auto_Start_Lector : Bool;
      Auto_Stop_Lector : Bool;
   END_VAR
   VAR
      State : UInt;
      R_Start_DB { S7_SetPoint := 'True'} : R_TRIG;
      T_Read_DB { S7_SetPoint := 'True'} : TON_TIME;
   END_VAR
   VAR_TEMP
      StartPos : Int;
      EndPos : Int;
      Code : String;
   END_VAR
BEGIN
   #R_Start_DB(CLK := #Station_Control.Start);

   IF #R_Start_DB.Q THEN
       IF #State = 0 THEN
           #State := 10;
       END_IF;
   END_IF;

   CASE #State OF
       0: // IDLE
           #Station_Control.Running := FALSE;
           #Station_Control.Ready := TRUE;
           #T_Read_DB(IN := FALSE,
                      PT := T#0S);

       10: // Start
           #Station_Control.Barcode := '';
           #Station_Control.Done := FALSE;
           #Station_Control.Valid := FALSE;
           #Station_Control.Ready := FALSE;
           #Station_Control.Running := TRUE;
           #State := 20;

       20: // Reading code
           #Station_Control.Start := FALSE;
           #Station_Control."Reading Gate number" := "FindStringField"(FieldName := 'Number', JsonStr := #Sick_Result);
           #Station_Control.Barcode := "FindStringField"(FieldName := 'Code', JsonStr := #Sick_Result);
           #Station_Control."Number of Reading Gates" := "FindStringField"(FieldName := 'NRG', JsonStr := #Sick_Result);
           #Auto_Start_Lector := TRUE;

           //Check if the gate is open
           IF #Station_Control."Number of Reading Gates" <> #Station_Control."Number of Reading Gates OLD" THEN
               #Station_Control."Number of Reading Gates OLD" := #Station_Control."Number of Reading Gates";
           END_IF;

           //Timer to read the barcode
           #T_Read_DB(IN := TRUE,
                      PT := T#15S);

           //If a new code was read or the time finished
           IF #Station_Control."Reading Gate number" <> #Station_Control."Reading Gate number OLD" OR #T_Read_DB.Q THEN
               #Auto_Start_Lector := FALSE; //Close the gate
               //New code
               IF #Station_Control."Reading Gate number" <> #Station_Control."Reading Gate number OLD" THEN
                   //Check if the string is not empty
                   IF LEN(IN := #Sick_Result) > 1 AND #Station_Control."Reading Gate number" <> '' THEN

                       // Find the start position of the code value
                       #StartPos := FIND(IN1 := #Sick_Result, IN2 := '"Code" :"');

                       IF #StartPos > 0 THEN

                           // Move to the first character of the code
                           #StartPos := #StartPos + LEN('"Code" :"');

                           // Find the next quotation mark after the code
                           #EndPos := FIND(
                                           IN1 := RIGHT(IN:=#Sick_Result, L:=LEN(#Sick_Result) - #StartPos + 1),
                                          IN2 := '"'
                           );

                           IF #EndPos > 0 THEN
                               #Code := MID(
                                            IN := #Sick_Result,
                                           L := #EndPos - 1,
                                           P := #StartPos
                               );
                           END_IF;

                       END_IF;
                       #Station_Control.Valid := TRUE;
                       #Station_Control.Barcode := #Code;
                       #Station_Control.Barcode_Old := #Station_Control.Barcode ;
                   ELSE //Empty
                       #Station_Control.Valid := FALSE;
                       #Station_Control.Barcode := '';
                   END_IF;
                   //Save OLD
                   #Station_Control."Reading Gate number OLD" := #Station_Control."Reading Gate number";
                   #T_Read_DB(IN := FALSE,
                              PT := T#0S);
                   #State := 30;
               ELSE // No code
                   #Station_Control.Valid := FALSE;
                   #Station_Control.Barcode := '';
                   #T_Read_DB(IN := FALSE,
                              PT := T#0S);
                   #State := 30;
               END_IF;
           END_IF;

       30: // Finally
           #Auto_Stop_Lector := TRUE; //Close gate
           //Make sure the command was sent
           IF #Auto_Stop_Lector THEN
               #Counter := #Counter + 1;
               #Station_Control.Running := FALSE;
               #Station_Control.Done := TRUE;
               #State := 0;
           END_IF;
   END_CASE;
END_FUNCTION_BLOCK

FUNCTION_BLOCK "Stack_Lights_FB"   // FB21, SCL
{ S7_Optimized_Access := 'TRUE' }
VERSION : 0.1
// stored: AutoNumber true, IsIECCheckEnabled false, IsRetainMemResEnabled false, MemoryReserve 100, SetENOAutomatically false, UDAEnableTagReadback false
   VAR_INPUT
      System_Auto : Bool;
      Fault : Bool;
   END_VAR
   VAR_OUTPUT
      Red : Bool;
      Green : Bool;
      Yellow : Bool;
   END_VAR
BEGIN
   //Commands for Stack Light

   IF #Fault THEN  // Fault = Red
       #Red := "Clock_0.5Hz";
       #Green := FALSE;
       #Yellow := FALSE;
   ELSIF #System_Auto THEN  // (1)Manual = Yellow
       #Yellow := FALSE;
       #Red := FALSE;
       #Green := TRUE;
   ELSIF NOT #System_Auto THEN  // (2)Semi-Auto = Blue
       #Green := FALSE;
       #Yellow := TRUE;
       #Red := FALSE;
   // ELSIF #System_Auto = 3 THEN  // (3)Auto = Green
   //     #Green := FALSE;
   //     #Red := FALSE;
   //     #Yellow := TRUE;

   ELSE
       #Green := FALSE;
       #Red := FALSE;
       #Yellow := FALSE;
   END_IF;
END_FUNCTION_BLOCK

FUNCTION_BLOCK "OPC_Control_FB"   // FB9, SCL
{ S7_Optimized_Access := 'TRUE' }
VERSION : 0.1
// stored: AutoNumber true, IsIECCheckEnabled false, IsRetainMemResEnabled false, MemoryReserve 100, SetENOAutomatically false, UDAEnableTagReadback false
   VAR_INPUT
      Id : UInt;
      All_In_Automatic : Bool;
      VTD_Error : Bool;
      OPC_Enable : Bool;
      Clear_OrderTable : Bool;
   END_VAR
   VAR_OUTPUT
      Error_ID : Word;
   END_VAR
   VAR
      Source_Location { ExternalAccessible := 'False'; ExternalVisible := 'False'; ExternalWritable := 'False'} : "ID_Decoded";
      Destination_Location { ExternalAccessible := 'False'; ExternalVisible := 'False'; ExternalWritable := 'False'} : "ID_Decoded";
      State_Main : UInt;
      State_VTD : UInt;
      State_Shuttle : UInt;
      State_CNV : UInt;
      T_Wait_Report_Done { S7_SetPoint := 'True'} : TON_TIME;
   END_VAR
   VAR_TEMP
      i : UInt;
      j : UInt;
      f : UInt;
      HMI_Reset : Bool;
   END_VAR
BEGIN
   IF "FirstScan" THEN
       "OPC_Enable" := TRUE;
   END_IF;

   REGION Errors STATE Main System
       IF #State_CNV > 0 AND #State_CNV < 250 THEN
           //CNV1
           IF #Source_Location.Device_Type = 10 OR #Destination_Location.Device_Type = 10 THEN
               IF "Control_DB".LCnv_Sys[#Id].Cnv_Level[#Source_Location.Level].Cnv1."Error"
                   OR
                   "Control_DB".LCnv_Sys[#Id].Cnv_Level[#Destination_Location.Level].Cnv1."Error" THEN
                   #Error_ID.%X3 := TRUE;
                   #State_CNV := 400;
               END_IF;
           END_IF;
           //CNV2
           IF #Source_Location.Device_Type = 11 OR #Destination_Location.Device_Type = 11 THEN
               IF "Control_DB".LCnv_Sys[#Id].Cnv_Level[#Source_Location.Level].Cnv2."Error"
                   OR
                   "Control_DB".LCnv_Sys[#Id].Cnv_Level[#Destination_Location.Level].Cnv2."Error" THEN
                   #Error_ID.%X3 := TRUE;
                   #State_CNV := 400;
               END_IF;
           END_IF;

           IF "Control_DB".ECnv_Sys[#Id].Error THEN
               #Error_ID.%X4 := TRUE;
               #State_CNV := 400;
           END_IF;
       END_IF;

       IF #State_VTD > 0 AND #State_VTD < 250 THEN
           IF #VTD_Error THEN
               #Error_ID.%X5 := TRUE;
               #State_VTD := 400;
           END_IF;
       END_IF;

       IF "Reset_All" THEN
           #Error_ID := 0;
       END_IF;
   END_REGION

   //Bit OPC in Error
   IF #State_VTD = 400 OR #State_Shuttle = 400 OR #State_CNV = 400 THEN
       #Error_ID.%X0 := TRUE;
   ELSE
       #Error_ID.%X0 := FALSE;
       #Error_ID.%X6 := FALSE;
       #Error_ID.%X7 := FALSE;
       #Error_ID.%X8 := FALSE;
   END_IF;

   IF ("Reset_All" OR #HMI_Reset) AND #State_VTD = 400
   THEN
       #State_VTD := 250;

   END_IF;

   IF ("Reset_All" OR #HMI_Reset) AND #State_Shuttle = 400
   THEN
       #State_Shuttle := 250;
   END_IF;

   IF ("Reset_All" OR #HMI_Reset) AND #State_CNV = 400
   THEN
       #State_CNV := 250;
   END_IF;

   (*
   Type of task to be performed:
       1 = Move to Floor
       2 = Shuttle Transfer into VTD
       3 = Shuttle Transfer out of VTD
       4 = Transfer Pallet into VTD
       5 = Transfer Pallet out of VTD
       6 = Transfer Pallet Roller to Roller
       7 = Transfer Pallet Chain to Chain  
       8 = Transfer to pick station 
       9 = Transfer from Pick station 
       10 = Weigh Pallet
       11 = Set chain Cnv as active (lower) // no use for now
       12 = Set Roller Cnv as active (raise) // no use for now

       Need to isolate ZZ in XXYYZZ to confirm #i = ZZ

       Extract XX (first two digits)
       xx := inputNumber / 10000;

       Extract YY (middle two digits)
       yy := (inputNumber / 100) MOD 100;

       Extract ZZ (last two digits)
       zz := inputNumber MOD 100;    
   *)


   IF #All_In_Automatic AND #OPC_Enable THEN
       REGION VTDs, Buffer conveyors and Shuttle 
           CASE #State_Main OF
               0:  //Pre operational state
                   #State_Main := 10;

               10: //Idle waiting for task
                   IF "Control_DB".WCS_OPC_Control[#Id].Task_Data_Available AND
                       #State_VTD = 0 AND #State_Shuttle = 0 AND #State_CNV = 0 THEN
                       #State_Main := 20;
                   END_IF;

               20: //Determine the type of task
                   "ID_Decode_F"(ID := "Control_DB".WCS_OPC_Control[#Id].Source_Location,
                                 ID_Decoded := #Source_Location);
                   "ID_Decode_F"(ID := "Control_DB".WCS_OPC_Control[#Id].Destination_Location,
                                 ID_Decoded := #Destination_Location);

                   //VTD move to floor
                   IF "Control_DB".WCS_OPC_Control[#Id].Task_Type = 1
                       AND NOT "Control_DB".VTD_Sys[#Id].Running THEN
                       #State_VTD := 30;
                       "Control_DB".WCS_OPC_Control[#Id].Task_Data_Available := 0;

                       //Shuttle transfer in/out of the VTD
                   ELSIF "Control_DB".WCS_OPC_Control[#Id].Task_Type = 2 OR "Control_DB".WCS_OPC_Control[#Id].Task_Type = 3
                   THEN
                       #State_Shuttle := 70;
                       "Control_DB".WCS_OPC_Control[#Id].Task_Data_Available := 0;

                       //Transfer Pallet in/out of the VTD
                   ELSIF ("Control_DB".WCS_OPC_Control[#Id].Task_Type = 4 OR "Control_DB".WCS_OPC_Control[#Id].Task_Type = 5)
                   THEN
                       #State_CNV := 100;
                       "Control_DB".WCS_OPC_Control[#Id].Task_Data_Available := 0;
                   END_IF;
           END_CASE;

           REGION VTD Move TO floor 
               CASE #State_VTD OF
                   0:  //Idle
                       ;

                   30: //Set all the Move to level variables
                       #State_Main := 0;
                       "Control_DB".VTD_Sys[#Id].Current_Task_Type := INT_TO_UINT("Control_DB".WCS_OPC_Control[#Id].Task_Type);
                       "Control_DB".VTD_Sys[#Id].Instruction.Pallet_Type := "Control_DB".WCS_OPC_Control[#Id].Pallet_Type;
                       "Control_DB".VTD_Sys[#Id].Instruction.Task_ID := INT_TO_UINT("Control_DB".WCS_OPC_Control[#Id].Task_ID);
                       "Control_DB".VTD_Sys[#Id].Instruction.Task_Metadata := "Control_DB".WCS_OPC_Control[#Id].Task_Metadata;
                       "Control_DB".VTD_Sys[#Id].Instruction.Move_To_Level := INT_TO_UINT(#Destination_Location.Level);
                       #State_VTD := 35;

                   // 35://Wait for the VTD to start its movement
                   //     "Control_DB".WCS_OPC_Control[#Id].SM_State := "Control_DB".VTD_Sys[#Id].SM_State;
                   //     IF "Control_DB".VTD_Sys[#Id].Enabled AND "Control_DB".VTD_Sys[#Id].Running THEN
                   //         "Control_DB".WCS_OPC_Control[#Id].Movement_Ready := TRUE;
                   //         #State_VTD := 40;
                   //     END_IF;

                   35://Wait for the VTD to start its movement
                       "Control_DB".WCS_OPC_Control[#Id].SM_State := "Control_DB".VTD_Sys[#Id].SM_State;
                       IF "Control_DB".VTD_Sys[#Id].Current_Level = #Destination_Location.Level THEN
                           //Already at destination level, skip movement
                           "Control_DB".WCS_OPC_Control[#Id].Movement_Ready := TRUE;
                           #State_VTD := 41;
                       ELSIF "Control_DB".VTD_Sys[#Id].Enabled AND "Control_DB".VTD_Sys[#Id].Running THEN
                           "Control_DB".WCS_OPC_Control[#Id].Movement_Ready := TRUE;
                           #State_VTD := 40;
                       END_IF;

                   40: //Wait for the VTD to complete its movement
                       "Control_DB".WCS_OPC_Control[#Id].SM_State := "Control_DB".VTD_Sys[#Id].SM_State;
                       IF "Control_DB".VTD_Sys[#Id].SM_State = 100 THEN
                           #State_VTD := 41;
                       END_IF;

                   41: //Wait for XXs for report done
                       #T_Wait_Report_Done.TON(IN := TRUE,
                                              PT := T#500ms);
                      IF #T_Wait_Report_Done.Q THEN
                          "Control_DB".WCS_OPC_Control[#Id].Movement_Request_Complete := TRUE;
                          #State_VTD := 45;
                      END_IF;

                   45: //Wait for the ACK before we go back to Idle
                       "Control_DB".WCS_OPC_Control[#Id].SM_State := "Control_DB".VTD_Sys[#Id].SM_State;
                       IF "Control_DB".WCS_OPC_Control[#Id].Movement_Request_Complete_Ack THEN///////////////////////////////////////////////////////////////////
                           #State_VTD := 250;
                       END_IF;

                   250: //Reset all variable and return to idle
                       "Control_DB".VTD_Sys[#Id].Instruction.Reset := FALSE;
                       "Control_DB".VTD_Sys[#Id].Instruction.Pallet_Type := 0;
                       "Control_DB".VTD_Sys[#Id].Instruction.Task_ID := 0;
                       "Control_DB".VTD_Sys[#Id].Instruction.Task_Metadata := '';
                       "Control_DB".VTD_Sys[#Id].Instruction.Move_To_Level := 0;
                       "Control_DB".VTD_Sys[#Id].Current_Task_Type := 0;

                       IF (#State_Shuttle = 0 OR #State_Shuttle = 250) AND
                           (#State_CNV = 0 OR #State_CNV = 250) THEN
                           //Reset the OPC control variables
                           "Control_DB".WCS_OPC_Control[#Id].SM_State := 0;
                           "Control_DB".WCS_OPC_Control[#Id].Movement_Ready := FALSE;
                           "Control_DB".WCS_OPC_Control[#Id].Movement_Request_Complete := FALSE;
                           "Control_DB".WCS_OPC_Control[#Id].Movement_Request_Complete_Ack := FALSE;
                           "Control_DB".WCS_OPC_Control[#Id].Pallet_Weight := 0;
                           "Control_DB".WCS_OPC_Control[#Id].Task_Metadata := '';
                           #T_Wait_Report_Done.TON(IN := FALSE,
                                                  PT := T#0S);
                          #State_VTD := 0;
                       END_IF;

                   400:// Error state
                       #Error_ID.%X6 := TRUE;
                       IF "Reset_All" OR #HMI_Reset
                       THEN
                           #Error_ID.%X5 := FALSE;
                           #Error_ID.%X6 := FALSE;
                           #State_VTD := 250;
                       END_IF;
               END_CASE;
           END_REGION ;

           REGION Transfer Shuttle in/out OF the VTD
               CASE #State_Shuttle OF
                   0:  //Idle
                       ;

                   70: //Set all the shuttle interlock variables
                       #State_Main := 0;
                       "Control_DB".VTD_Sys[#Id].Instruction.Task_ID := "Control_DB".WCS_OPC_Control[#Id].Task_ID; //Assign task ID to WCS Task ID
                       "Control_DB".VTD_Sys[#Id].Instruction.Task_Metadata := "Control_DB".WCS_OPC_Control[#Id].Task_Metadata;
                       "Control_DB".VTD_Sys[#Id].Instruction.Pallet_Type := "Control_DB".WCS_OPC_Control[#Id].Pallet_Type;
                       "Control_DB".VTD_Sys[#Id].Current_Task_Type := INT_TO_UINT("Control_DB".WCS_OPC_Control[#Id].Task_Type);
                       "Control_DB".VTD_Sys[#Id].Shuttle_Interlock.Shuttle_Interlock_Task_ID := INT_TO_UINT("Control_DB".WCS_OPC_Control[#Id].Task_ID);
                       "Control_DB".VTD_Sys[#Id].Shuttle_Interlock.Shuttle_Interlock_Task_Metadata := "Control_DB".WCS_OPC_Control[#Id].Task_Metadata;
                       "Control_DB".VTD_Sys[#Id].Shuttle_Interlock.Shuttle_ID := INT_TO_UINT("Control_DB".WCS_OPC_Control[#Id].Shuttle_ID);
                       "Control_DB".VTD_Sys[#Id].Shuttle_Interlock.Shuttle_Loaded := "Control_DB".WCS_OPC_Control[#Id].Shuttle_Loaded;
                       "Control_DB".VTD_Sys[#Id].Shuttle_Interlock.Shuttle_Start_Location := "Control_DB".WCS_OPC_Control[#Id].Source_Location;
                       "Control_DB".VTD_Sys[#Id].Shuttle_Interlock.Shuttle_Target_Location := "Control_DB".WCS_OPC_Control[#Id].Destination_Location;

                       "Control_DB".VTD_Sys[#Id].Shuttle_Interlock.Interlock_Request := TRUE;
                       #State_Shuttle := 75;

                   75: //Inform WCS that the VTD is ready to interlock
                       "Control_DB".WCS_OPC_Control[#Id].SM_State := "Control_DB".VTD_Sys[#Id].SM_State;
                       IF "Control_DB".VTD_Sys[#Id].Shuttle_Interlock.Ready_To_Interlock THEN
                           "Control_DB".WCS_OPC_Control[#Id].Movement_Ready := TRUE;
                           "Control_DB".WCS_OPC_Control[#Id].Task_Data_Available := FALSE;
                           #State_Shuttle := 80;
                       END_IF;

                   80://Inform WCS that the interlock is complete
                       IF "Control_DB".VTD_Sys[#Id].Shuttle_Interlock.Interlock_Complete THEN
                           "Control_DB".VTD_Sys[#Id].Shuttle_Interlock.Interlock_Request := FALSE;
                           "Control_DB".WCS_OPC_Control[#Id].Movement_Request_Complete := TRUE;
                           #State_Shuttle := 90;
                       END_IF;

                       // 81: //Wait for XXs for report done
                   //     #T_Wait_Report_Done.TON(IN := TRUE,
                   //                            PT := T#500mS);
                   //    IF #T_Wait_Report_Done.Q THEN
                   //         #State_Shuttle := 90;
                   //     END_IF;

                   90: //Reset VTD back to idle state
                       IF "Control_DB".WCS_OPC_Control[#Id].Movement_Request_Complete_Ack THEN
                           "Control_DB".VTD_Sys[#Id].Shuttle_Interlock.Interlock_Complete_Ack := TRUE;
                           #State_Shuttle := 250;
                       END_IF;

                   250: //Reset all variable and return to idle
                       //Reset Shuttle interlock
                       "Control_DB".VTD_Sys[#Id].Shuttle_Interlock.Interlock_Request := FALSE;
                       "Control_DB".VTD_Sys[#Id].Shuttle_Interlock.Shuttle_Start_Location := 0;
                       "Control_DB".VTD_Sys[#Id].Shuttle_Interlock.Shuttle_Target_Location := 0;
                       "Control_DB".VTD_Sys[#Id].Shuttle_Interlock.Shuttle_Loaded := 0;
                       "Control_DB".VTD_Sys[#Id].Shuttle_Interlock.Shuttle_ID := 0;
                       "Control_DB".VTD_Sys[#Id].Shuttle_Interlock.Shuttle_Interlock_Task_ID := 0;
                       "Control_DB".VTD_Sys[#Id].Shuttle_Interlock.Shuttle_Interlock_Task_Metadata := '';
                       "Control_DB".VTD_Sys[#Id].Shuttle_Interlock.Interlock_Complete_Ack := FALSE;

                       IF (#State_VTD = 0 OR #State_VTD = 250) AND
                           (#State_CNV = 0 OR #State_CNV = 250) THEN
                           //Reset the OPC control variables
                           "Control_DB".WCS_OPC_Control[#Id].SM_State := 0;
                           "Control_DB".WCS_OPC_Control[#Id].Movement_Ready := FALSE;
                           "Control_DB".WCS_OPC_Control[#Id].Movement_Request_Complete := FALSE;
                           "Control_DB".WCS_OPC_Control[#Id].Movement_Request_Complete_Ack := FALSE;
                           "Control_DB".WCS_OPC_Control[#Id].Task_Metadata := '';
                           #T_Wait_Report_Done.TON(IN := FALSE,
                                                  PT := T#0S);

                           #State_Shuttle := 0;
                       END_IF;

                   400:// Error state
                       #Error_ID.%X7 := TRUE;
                       IF "Reset_All" OR #HMI_Reset
                       THEN
                           #Error_ID.%X7 := FALSE;
                           #State_Shuttle := 250;
                       END_IF;
               END_CASE;
           END_REGION ;

           REGION Transfer Pallet in/out OF the VTD
               CASE #State_CNV OF
                   0:  //Idle
                       ;

                   100: //Set the destination conveyor variables
                       #State_Main := 0;

                       //Assign task to receiving conveyor
                       IF #Destination_Location.Level >= "Settings_DB".VTD_Sys[#Id].Lowest_Level AND #Destination_Location.Level <= "Settings_DB".VTD_Sys[#Id].Highest_Level THEN

                           //Buffer conveyors
                           //CNV 1
                           IF (#Destination_Location.Device_Type = 10 AND "Control_DB".ECnv_Sys[#Id].Cnv_Occupied AND
                               NOT "Control_DB".LCnv_Sys[#Id].Cnv_Level[#Destination_Location.Level].Cnv1.Cnv_Occupied) OR
                               (#Destination_Location.Device_Type = 10 AND #Destination_Location.Level = 1 AND #Source_Location.Device_Type = 0 AND
                               NOT "Control_DB".LCnv_Sys[#Id].Cnv_Level[#Destination_Location.Level].Cnv1.Cnv_Occupied)
                           THEN
                               "Control_DB".LCnv_Sys[#Id].Cnv_Level[#Destination_Location.Level].Cnv1.Instruction.Task_ID := INT_TO_UINT("Control_DB".WCS_OPC_Control[#Id].Task_ID);
                               "Control_DB".LCnv_Sys[#Id].Cnv_Level[#Destination_Location.Level].Cnv1.Instruction.Task_Metadata := "Control_DB".WCS_OPC_Control[#Id].Task_Metadata;
                               "Control_DB".LCnv_Sys[#Id].Cnv_Level[#Destination_Location.Level].Cnv1.Current_Task_Type := INT_TO_UINT("Control_DB".WCS_OPC_Control[#Id].Task_Type);
                               "Control_DB".LCnv_Sys[#Id].Cnv_Level[#Destination_Location.Level].Cnv1.Instruction.Transfer_From_ID := "Control_DB".WCS_OPC_Control[#Id].Source_Location;
                               "Control_DB".LCnv_Sys[#Id].Cnv_Level[#Destination_Location.Level].Cnv1.Instruction.Transfer_To_ID := "Control_DB".WCS_OPC_Control[#Id].Destination_Location;
                               IF "Control_DB".WCS_OPC_Control[#Id].Pallet_Type = 'E' AND "Control_DB".WCS_OPC_Control[#Id].Pallet_Alignment = 'L' THEN
                                   "Control_DB".LCnv_Sys[#Id].Cnv_Level[#Destination_Location.Level].Cnv1.Instruction.Pallet_Type := 3;
                               ELSIF "Control_DB".WCS_OPC_Control[#Id].Pallet_Type = 'E' AND "Control_DB".WCS_OPC_Control[#Id].Pallet_Alignment = 'R' THEN
                                   "Control_DB".LCnv_Sys[#Id].Cnv_Level[#Destination_Location.Level].Cnv1.Instruction.Pallet_Type := 2;
                               END_IF;

                               //Enable the conveyor and start the transfer
                               "Control_DB".LCnv_Sys[#Id].Cnv_Level[#Destination_Location.Level].Cnv1.Instruction.Start_Transfer := TRUE;
                               #State_CNV := 105;

                               //CNV 2
                           ELSIF #Destination_Location.Device_Type = 11 AND "Control_DB".ECnv_Sys[#Id].Cnv_Occupied AND
                               NOT "Control_DB".LCnv_Sys[#Id].Cnv_Level[#Destination_Location.Level].Cnv2.Cnv_Occupied
                           THEN
                               "Control_DB".LCnv_Sys[#Id].Cnv_Level[#Destination_Location.Level].Cnv2.Instruction.Task_ID := INT_TO_UINT("Control_DB".WCS_OPC_Control[#Id].Task_ID);
                               "Control_DB".LCnv_Sys[#Id].Cnv_Level[#Destination_Location.Level].Cnv2.Instruction.Task_Metadata := "Control_DB".WCS_OPC_Control[#Id].Task_Metadata;
                               "Control_DB".LCnv_Sys[#Id].Cnv_Level[#Destination_Location.Level].Cnv2.Current_Task_Type := INT_TO_UINT("Control_DB".WCS_OPC_Control[#Id].Task_Type);
                               "Control_DB".LCnv_Sys[#Id].Cnv_Level[#Destination_Location.Level].Cnv2.Instruction.Transfer_From_ID := "Control_DB".WCS_OPC_Control[#Id].Source_Location;
                               "Control_DB".LCnv_Sys[#Id].Cnv_Level[#Destination_Location.Level].Cnv2.Instruction.Transfer_To_ID := "Control_DB".WCS_OPC_Control[#Id].Destination_Location;
                               IF "Control_DB".WCS_OPC_Control[#Id].Pallet_Type = 'E' AND "Control_DB".WCS_OPC_Control[#Id].Pallet_Alignment = 'L' THEN
                                   "Control_DB".LCnv_Sys[#Id].Cnv_Level[#Destination_Location.Level].Cnv2.Instruction.Pallet_Type := 3;
                               ELSIF "Control_DB".WCS_OPC_Control[#Id].Pallet_Type = 'E' AND "Control_DB".WCS_OPC_Control[#Id].Pallet_Alignment = 'R' THEN
                                   "Control_DB".LCnv_Sys[#Id].Cnv_Level[#Destination_Location.Level].Cnv2.Instruction.Pallet_Type := 2;
                               END_IF;

                               //Enable the conveyor and start the transfer
                               "Control_DB".LCnv_Sys[#Id].Cnv_Level[#Destination_Location.Level].Cnv2.Instruction.Start_Transfer := TRUE;
                               #State_CNV := 105;

